(* IEC 61131-3 sources: daoli-st-library/DL_Process (part 45) *)

(* ---- FB_DL_PileClampCtrl.st ---- *)
(*
  FB_DL_PileClampCtrl  —  堆叠压紧板两段压力-位移控制 / Pile clamp two-stage pressure-position control
  分类 Category : DL_Process
  码位 Code     : 16#06_0_90
  版本 Version  : 1.0.0
  溯源 Source   : LBP（Lediberg Process Library）语义借鉴 · clean-room 实现，仅借分类/参数域/命名，未复制源码
  功能 Function : 1) 压紧板「预压 → 全压」两段顺控（复用 FB_DL_StepSequencer 推步 + I_DL_Cylinder 缸接口依赖注入）；
                  2) 预压段压力-位移落窗才放行全压段（禁跳段）；
                  3) 保压计时独立 TON 且 IN := NOT ton.Q 自复位（FB33-2）。
  边界 Boundary : ① 预压未达窗禁进全压段（步完成信号由本件门控）；
                  ② 压力/位移任一无效：冻结当前段并保持命令（不追加新指令）；
                  ③ 包络窗口上下限倒置出厂报码不运行；
                  ④ 释压命令与压紧命令互斥，同拍双真取释压（安全侧）；
                  ⑤ 输出三行同向：缸命令 → 段状态 → 完成标志。
  依赖 Depends  : FB_DL_StepSequencer（两段推步，每拍无条件调用）
                  I_DL_Cylinder（缸接口，VAR_IN_OUT 引用注入，引用非空判零 (ipCyl <> 0) 门控）

  码表 Error codes（本件子码步进 16#30 · 本格 90 与既有 9X 子码段冲突，错位至 C0/D0 避让）:
    16#0002_06C0 故障级：组态非法（两段目标倒置 / 包络窗倒置 / 保压时长 <= 0）
    16#0002_06D0 故障级：步超时（段内压力-位移未在限时内落窗，映射自顺控实例）
    16#0002_06B0 信息级：压力或位移无效当前段冻结（不置 bError）
*)

TYPE E_DL_PccPhase :
(
    eIdle    := 0,   // 空闲 / Idle
    ePre     := 10,  // 预压段 / Pre-clamp stage
    eFull    := 20,  // 全压段 / Full-clamp stage
    eHold    := 30,  // 保压段 / Pressure holding
    eRelease := 40,  // 释压段 / Release stage
    eDone    := 50,  // 压紧完成 / Clamp done
    eFrozen  := 60,  // 反馈无效冻结 / Frozen by invalid feedback
    eFault   := 90   // 故障锁定 / Fault locked
);
END_TYPE

FUNCTION_BLOCK FB_DL_PileClampCtrl
VAR_INPUT
    bClampReq     : BOOL;                           // 压紧命令（电平）/ Clamp command, level
    bReleaseReq   : BOOL;                           // 释压命令（电平，与压紧互斥取优先）/ Release command, level
    bReset        : BOOL;                           // 复位，上升沿清故障 / Reset, clears fault
    fPressKN      : REAL;                           // 压紧压力实测 [kN] / Measured clamp pressure [kN]
    fPosMm        : REAL;                           // 压紧板位移实测 [mm] / Measured plate position [mm]
    fPreTargetKN  : REAL := 5.0;                    // 预压段目标压力 [kN] / Pre-stage target pressure [kN]
    fFullTargetKN : REAL := 12.0;                   // 全压段目标压力 [kN] / Full-stage target pressure [kN]
    fPreWinKN     : REAL := 0.8;                    // 预压窗半宽 [kN]，域 > 0 / Pre-stage window half width [kN]
    fFullWinKN    : REAL := 1.0;                    // 全压窗半宽 [kN]，域 > 0 / Full-stage window half width [kN]
    fPrePosLoMm   : REAL := 3.0;                    // 预压段位移窗下限 [mm] / Pre-stage position window low [mm]
    fPrePosHiMm   : REAL := 6.0;                    // 预压段位移窗上限 [mm] / Pre-stage position window high [mm]
    fFullPosLoMm  : REAL := 7.5;                    // 全压段位移窗下限 [mm] / Full-stage position window low [mm]
    fFullPosHiMm  : REAL := 10.0;                   // 全压段位移窗上限 [mm] / Full-stage position window high [mm]
    tHoldTime     : TIME := T#5S;                   // 保压时长 [s]，域 > 0 / Holding duration
    fEps          : REAL := 1.0E-6;                 // 浮点判零容差 [1] / Floating zero tolerance
END_VAR
VAR_IN_OUT
    ipCyl         : I_DL_Cylinder;                  // 压紧缸接口（依赖注入）/ Clamp cylinder interface, injected
END_VAR
VAR_OUTPUT
    bClampCmd     : BOOL;                           // 缸压紧命令出口 / Cylinder clamp command output
    bReleaseCmd   : BOOL;                           // 缸释压命令出口 / Cylinder release command output
    eStageOut     : E_DL_PccPhase;                  // 当前段状态 / Current stage status
    bClampDone    : BOOL;                           // 压紧完成标志（保持型）/ Clamp done flag, held
    bEnvViol      : BOOL;                           // 包络越窗标志（本拍重算）/ Envelope violation flag
    bError        : BOOL;                           // 故障标志，与故障级码配对 / Fault flag
    uErrorId      : UDINT;                          // 事件码，0 = 无事件 / Event code
END_VAR
VAR
    fbSeq         : FB_DL_StepSequencer;            // 两段顺控实例（无条件调用）/ Two-step sequencer instance
    rtrReset      : R_TRIG;                         // 复位沿 / Reset edge
    tonHold       : TON;                            // 保压计时器（IN := NOT Q 自复位范式不适用本件：保压为单次电平计时）/ Holding timer
    abStepDone    : ARRAY[0..15] OF BOOL;           // 步完成信号表 / Step-done table
    auStepTo      : ARRAY[0..15] OF TIME;           // 步超时表 / Step timeout table
    _eState       : E_DL_PccPhase := E_DL_PccPhase.eIdle;  // 内部状态 / Internal state
    bCfgOk        : BOOL;                           // 组态合法标志 / Configuration valid
    bRefOk        : BOOL;                           // 缸接口引用有效 / Interface reference valid
    bFbOk         : BOOL;                           // 压力/位移双有效 / Pressure and position valid
    bPreInWin     : BOOL;                           // 预压段压力-位移落窗 / Pre-stage in window
    bFullInWin    : BOOL;                           // 全压段压力-位移落窗 / Full-stage in window
    bHoldDone     : BOOL;                           // 保压计时到 / Holding time elapsed
    uFault        : UDINT;                          // 锁存故障码 / Latched fault code
    uInfo         : UDINT;                          // 信息级码 / Information code
END_VAR

(* === 段 0 · 实例刷新 === *)
rtrReset(CLK := bReset);                          // 每拍刷新复位沿

(* === 段 1 · 组态闸与反馈域闸 === *)
bRefOk := (ipCyl <> 0);                           // 接口引用有效性（引用非空判零口径，R4 防御）/ Interface reference validity, null-reference test
bCfgOk := (fFullTargetKN > fPreTargetKN + fEps)   // 两段目标不倒置（全压 > 预压）
          AND (fPreWinKN > fEps) AND (fFullWinKN > fEps)
          AND (fPrePosHiMm > fPrePosLoMm + fEps)  // 预压位移窗不倒置
          AND (fFullPosHiMm > fFullPosLoMm + fEps)// 全压位移窗不倒置
          AND (TIME_TO_REAL(tHoldTime) > fEps)    // 保压时长正域
          AND (fPreTargetKN = fPreTargetKN) AND (fFullTargetKN = fFullTargetKN);  // NaN 自反
IF NOT bCfgOk THEN
    uFault := 16#0002_06C0;                       // 故障级：组态非法
END_IF
IF rtrReset.Q AND bCfgOk THEN
    uFault := 16#0000;                            // 复位沿清锁存（解除路径可达）
END_IF
uInfo := 16#0000;                                 // 信息码每拍清零
bFbOk := (fPressKN = fPressKN) AND (ABS(fPressKN) < 1.0E30)
         AND (fPosMm = fPosMm) AND (ABS(fPosMm) < 1.0E30);      // 双反馈 NaN 自反 + 幅值闸
IF NOT bFbOk THEN
    uInfo := 16#0002_06B0;                        // 信息级：反馈无效当前段冻结
END_IF

(* === 段 2 · 窗口判定（本拍重算）=== *)
bPreInWin := bFbOk AND (ABS(fPressKN - fPreTargetKN) <= fPreWinKN + fEps)
             AND (fPosMm >= fPrePosLoMm - fEps) AND (fPosMm <= fPrePosHiMm + fEps);   // 预压落窗
bFullInWin := bFbOk AND (ABS(fPressKN - fFullTargetKN) <= fFullWinKN + fEps)
              AND (fPosMm >= fFullPosLoMm - fEps) AND (fPosMm <= fFullPosHiMm + fEps);  // 全压落窗
bEnvViol := bFbOk AND (fPressKN > fFullTargetKN + fFullWinKN + 5.0 * fFullWinKN);   // 包络越窗：压力远超全压窗

(* === 段 3 · 顺控实例装载（每拍无条件调用）=== *)
abStepDone[0] := bPreInWin;                       // 步 0 = 预压：落窗才算完成（门控禁跳段）
abStepDone[1] := bFullInWin;                      // 步 1 = 全压：落窗才算完成
abStepDone[2] := TRUE;                            // 步 2 = 保压：完成由本件 TON 判
auStepTo[0] := T#30S;                             // 预压步超时 30 s
auStepTo[1] := T#30S;                             // 全压步超时 30 s
auStepTo[2] := T#0S;                              // 保压步不监控（由保压 TON 承担）
fbSeq(bStart := bClampReq AND (NOT bReleaseReq) AND bCfgOk AND bRefOk AND bFbOk,   // 压紧命令且非释压优先
      abStepDone := abStepDone,                   // 步完成表
      auStepTimeout := auStepTo,                  // 步超时表
      bHold := NOT bFbOk,                         // 反馈无效：顺控保持（冻结当前段）
      bAbort := bReleaseReq OR (NOT bCfgOk),      // 释压/组态故障：中止回空闲
      bReset := rtrReset.Q);                      // 复位沿透传
IF fbSeq.bError THEN
    uFault := 16#0002_06D0;                       // 故障级：步超时（映射自顺控实例）
END_IF

(* === 段 4 · 保压计时（独立 TON，段内电平触发）=== *)
bHoldDone := FALSE;                               // 保压完成本拍重算
IF fbSeq.nCurrentStep = 2 THEN                    // 顺控进入保压步才计时
    tonHold(IN := TRUE, PT := tHoldTime);         // 保压计时（步号门控自清，离开步 IN 即断）
    IF tonHold.Q THEN
        bHoldDone := TRUE;                        // 保压时长到
    END_IF
ELSE
    tonHold(IN := FALSE, PT := tHoldTime);        // 离开保压步：定时器断输入复位（R40 分段监控按段断输入）
END_IF

(* === 段 5 · 主状态机（ENUM + CASE，含 ELSE 兜底）=== *)
CASE _eState OF
E_DL_PccPhase.eIdle :
    bClampDone := FALSE;                          // 空闲未完成
    IF uFault <> 16#0000 THEN
        _eState := E_DL_PccPhase.eFault;          // 故障优先
    END_IF
    IF fbSeq.bRunning AND (fbSeq.nCurrentStep = 0) THEN
        _eState := E_DL_PccPhase.ePre;            // 顺控步 0：预压相
    END_IF

E_DL_PccPhase.ePre :
    IF fbSeq.nCurrentStep = 1 THEN
        _eState := E_DL_PccPhase.eFull;           // 步 1：全压相（预压未落窗顺控不推步）
    ELSIF fbSeq.nCurrentStep < 0 THEN
        _eState := E_DL_PccPhase.eIdle;           // 顺控中止回空闲
    END_IF

E_DL_PccPhase.eFull :
    IF fbSeq.nCurrentStep = 2 THEN
        _eState := E_DL_PccPhase.eHold;           // 步 2：保压相
    ELSIF fbSeq.nCurrentStep < 0 THEN
        _eState := E_DL_PccPhase.eIdle;           // 顺控中止回空闲
    END_IF

E_DL_PccPhase.eHold :
    IF bHoldDone THEN
        _eState := E_DL_PccPhase.eDone;           // 保压满：完成相
    ELSIF bReleaseReq THEN
        _eState := E_DL_PccPhase.eRelease;        // 释压优先（安全侧同拍双真取释压）
    END_IF

E_DL_PccPhase.eRelease :
    IF fbSeq.nCurrentStep < 0 THEN
        _eState := E_DL_PccPhase.eIdle;           // 释压完成回空闲（解除路径可达）
    END_IF

E_DL_PccPhase.eDone :
    bClampDone := TRUE;                           // 完成保持（防同拍抹除）
    IF bReleaseReq OR (NOT bClampReq) THEN
        bClampDone := FALSE;                      // 释压或撤命令：完成复位
        _eState := E_DL_PccPhase.eIdle;           // 回空闲
    END_IF

E_DL_PccPhase.eFrozen :
    IF bFbOk THEN
        _eState := E_DL_PccPhase.ePre;            // 反馈恢复回预压相续判（解除路径可达）
    END_IF

E_DL_PccPhase.eFault :
    IF uFault = 16#0000 THEN
        _eState := E_DL_PccPhase.eIdle;           // 解锁回空闲
    END_IF

ELSE
    _eState := E_DL_PccPhase.eFault;              // 非法状态拦截
    uFault := 16#0002_06C0;                       // 故障级：相 ID 越界复用组态码段
END_CASE
IF (NOT bFbOk) AND (_eState = E_DL_PccPhase.ePre OR _eState = E_DL_PccPhase.eFull
    OR _eState = E_DL_PccPhase.eHold) THEN
    _eState := E_DL_PccPhase.eFrozen;             // 运行段中反馈丢失：转冻结相（命令保持）
END_IF

(* === 段 6 · 缸命令出口映射（互斥：释压优先）=== *)
bClampCmd := (_eState = E_DL_PccPhase.ePre) OR (_eState = E_DL_PccPhase.eFull)
             OR (_eState = E_DL_PccPhase.eHold);  // 压紧命令只在压紧段保持
bClampCmd := bClampCmd AND bFbOk AND bRefOk AND (uFault = 16#0000);   // 无效/故障安全侧撤命令
bReleaseCmd := (_eState = E_DL_PccPhase.eRelease) OR bReleaseReq;     // 释压命令（同拍双真取释压）
bReleaseCmd := bReleaseCmd AND bRefOk;            // 引用无效不出命令
IF bRefOk AND bReleaseCmd THEN
    ipCyl.CmdRetract();                           // 释压指令（接口依赖注入调用）
ELSIF bRefOk AND bClampCmd THEN
    ipCyl.CmdExtend();                            // 压紧指令（接口依赖注入调用）
END_IF

(* === 段 7 · 输出映射 === *)
bError := (uFault <> 16#0000);                    // 故障标志仅由故障级码置位（R45 配对）
IF bError THEN
    uErrorId := uFault;                           // 故障级优先上报
ELSE
    uErrorId := uInfo;                            // 否则上报信息级码
END_IF
eStageOut := _eState;                             // 输出枚举段尾单点映射（N2 规则）
END_FUNCTION_BLOCK

(* ---- FB_DL_PilePressLimitClass.st ---- *)
(*
  Component : FB_DL_PilePressLimitClass
  Category  : DL_Process
  Type      : FB
  Version   : 1.0.0
  CodeSeg   : 16#06_0_3A
  Summary   : 堆叠压力四档分级与 NG 分道：压力归类（A/B/C/NG 四档，档界常量带单位）+ 分道放行。
              Stacking pressure four-band classification and NG routing: band classify with unit-tagged limits plus lane release.
  溯源声明  : 参照 FC_DL_LimitClassify 语义（clean-room 自含实现，无实例依赖）
  边界安全  : 压力非有限（NaN 自反 + Inf 上限）与负值域拦截（kN）；档界常量域闸（L1 < L2 < L3，
              防档位倒置）；判定电平比较（非等值直比）；分道放行带起动沿防重复放行；
              各档计数独立且防回卷；全浮点比较带 fEps 容差。
  复用      : 参照 FC_DL_LimitClassify 语义（clean-room 自含实现，无实例依赖）
*)

FUNCTION_BLOCK FB_DL_PilePressLimitClass
VAR_INPUT
    bRun     : BOOL;                    (* 分级使能 · Enable *)
    fPressKN : LREAL;                   (* 堆叠压力 [kN] · Stacking pressure *)
    bPiecePulse: BOOL;                  (* 单件到位脉冲 [事件] · Piece-in-place pulse *)
    fL1KN    : LREAL := 8.0;            (* A 档下界 [kN] · Band A lower bound *)
    fL2KN    : LREAL := 6.0;            (* B 档下界 [kN] · Band B lower bound *)
    fL3KN    : LREAL := 4.0;            (* C 档下界 [kN] · Band C lower bound *)
    fEps     : LREAL := 1.0E-6;         (* 浮点判零容差 [实数域] · Floating zero tolerance *)
END_VAR
VAR_OUTPUT
    eClass   : (eClsA := 0, eClsB := 1, eClsC := 2, eClsNG := 3);   (* 档位枚举输出 / Class output enum *)
    bNgLane  : BOOL;                    (* NG 分道放行 [引脚] · NG lane release *)
    bOkLane  : BOOL;                    (* 合格道放行 [引脚] · OK lane release *)
    nCntA    : UDINT;                   (* A 档累计 [件]，防回卷 · Band A count *)
    nCntB    : UDINT;                   (* B 档累计 [件]，防回卷 · Band B count *)
    nCntC    : UDINT;                   (* C 档累计 [件]，防回卷 · Band C count *)
    nCntNG   : UDINT;                   (* NG 档累计 [件]，防回卷 · NG count *)
    bError   : BOOL;                    (* 故障标志，与故障码配对 · Fault flag paired with codes *)
    uErrorId : UDINT;                   (* 事件码 16#0000_003A，0 无事件 · Event code *)
END_VAR
VAR
    uCode    : WORD;    (* 码位暂存，每拍重算 [码] · Code staging *)
    bSigOk   : BOOL;    (* 输入有效标志 · Input validity flag *)
    bThrOk   : BOOL;    (* 档界整定域标志 · Band limit tuning validity *)
    bPiecePrv: BOOL;    (* 上拍到位脉冲快照，上升沿判据 · Previous pulse snapshot *)
    bPiece   : BOOL;    (* 到位上升沿 [脉冲] · Piece rising edge *)
    bClassNow: BOOL;    (* 本拍已归类标志（防重复放行）/ Classified this scan *)
    nCycles  : UDINT;   (* 有效归类拍计数 [拍]，防回卷 · Classify scan count *)
END_VAR
VAR CONSTANT
    DL_PLC_WRAP : UDINT := 4294967290;  (* 计数防回卷余量 [件] · Counter wrap guard *)
END_VAR

(* === 段 0 · 实例刷新 === *)
(* 无 TON/R_TRIG 实例：沿判据用快照实现；No timer instances, edges via snapshots *)
bPiece := bPiecePulse AND (NOT bPiecePrv);      (* 到位上升沿 / Piece rising edge *)
bPiecePrv := bPiecePulse;                       (* 快照更新 / Snapshot *)

(* === 段 1 · 输入校验与量程闸 === *)
uCode := 16#0000;                       // 每拍清码（可达清零基线）/ Clear codes each scan
bSigOk := (fPressKN = fPressKN) AND (ABS(fPressKN) < 1.0E308)   // 非有限拦截 / Non-finite guard
          AND (fPressKN >= 0.0);                                        // 压力非负域闸 / Non-negative pressure
bThrOk := (fL3KN > fEps) AND (fL2KN > fL3KN) AND (fL1KN > fL2KN);   // 档界倒置闸（L1>L2>L3）/ Band order gate
IF NOT bSigOk OR NOT bThrOk THEN
    uCode := 16#003A;                   // 故障级：域外或档界倒置 / Fault: domain or band order invalid
END_IF

(* === 段 2 · 主逻辑：四档归类与分道放行 === *)
bOkLane := FALSE;                       (* 放行输出为脉冲量，默认收口 / Lane outputs are pulses *)
bNgLane := FALSE;
IF bSigOk AND bThrOk THEN
    IF bPiece THEN                      (* 到位沿：归类一次 / Classify once on the edge *)
        bClassNow := TRUE;              (* 本拍已归类 / Classified *)
        IF fPressKN >= fL1KN THEN
            eClass := eClsA;            (* A 档（输出枚举在沿上直赋，非 CASE 状态机）/ Band A *)
            IF nCntA < DL_PLC_WRAP THEN
                nCntA := nCntA + 1;     (* A 档计数 / Count band A *)
            END_IF
            bOkLane := TRUE;            (* 合格道放行 / Release the OK lane *)
        ELSIF fPressKN >= fL2KN THEN
            eClass := eClsB;            (* B 档 / Band B *)
            IF nCntB < DL_PLC_WRAP THEN
                nCntB := nCntB + 1;
            END_IF
            bOkLane := TRUE;
        ELSIF fPressKN >= fL3KN THEN
            eClass := eClsC;            (* C 档 / Band C *)
            IF nCntC < DL_PLC_WRAP THEN
                nCntC := nCntC + 1;
            END_IF
            bOkLane := TRUE;
        ELSE
            eClass := eClsNG;           (* NG 档：低于 C 下界 / NG below the C bound *)
            IF nCntNG < DL_PLC_WRAP THEN
                nCntNG := nCntNG + 1;
            END_IF
            bNgLane := TRUE;            (* NG 分道放行 / Release the NG lane *)
        END_IF
        IF nCycles < DL_PLC_WRAP THEN
            nCycles := nCycles + 1;     (* 归类拍计数 / Count classifications *)
        END_IF
    END_IF
END_IF

(* === 段 3 · 输出映射与故障码 === *)
IF NOT (bPiece OR bClassNow) THEN
    (* 非归类拍保持上次档位输出（回放语义）/ Keep the last class between pieces *)
END_IF
IF NOT bRun THEN
    bClassNow := FALSE;                 (* 撤使能清归类态（可达复位）/ Clear on disable *)
    bOkLane := FALSE;
    bNgLane := FALSE;
END_IF
bError := (uCode <> 16#0000);           (* 故障标志配对 / Fault flag paired *)
uErrorId := WORD_TO_UDINT(uCode);       (* 码位单点写入（16#0000_003A 形态）/ Single write point *)
END_FUNCTION_BLOCK

(* ---- FB_DL_PipeScannerRoute.st ---- *)
(*
  FB_DL_PipeScannerRoute  —  管输批次扫码分输（扫码枪契约 + 阀序分道） / Pipe batch scan-and-route: scanner contract plus valve sequence routing
  分类 Category : DL_Process
  版本 Version  : 1.0.0
  来源 Source   : t2-2-lbp — 管输分输族深化
  溯源 Origin   : clean-room 实现，未复制任何源码行
  功能 Function : 1) 四相顺控：eIdle（等批次到达沿）→ eWaitScan（等扫码枪契约
                  bScanValid，tScanTo 超时判）→ eValve（按 uBatchId MOD nRoutes
                  分道，开阀等阀位反馈）→ eDone（关阀回 eIdle）；
                  2) 扫码契约：uBatchId 仅在 bScanValid 当拍采信（锁存快照），
                  分道号 nRouteIdx := UDINT_TO_DINT(uBatchId MOD nRoutes)
                  （模基数域闸 1..4，无除零）；
                  3) 故障级：0388 组态非法（分道数越域）+ ELSE 兜底归并 /
                  0389 扫码缺失超窗锁存 / 038A 开阀后阀位反馈不一致锁存；
                  4) 信息级三码：扫码成功 / 分道指令发出 / 分道完成（单拍沿）；
                  5) 解除式全当拍量（R240 落地），逐 BOOL 标注见段 4。
  边界 Boundary : ① 超时 TON 均单相独占（IN 为单相等式），跨相迁移拍 IN 必断
                  （R228-A）；阀超时与扫码超时分实例；
                  ② 阀反馈判据仅认当拍量 a_bValveFb，禁锁存反馈自指；
                  ③ 分道索引域 0..3 由 nRoutes 域闸 1..4 与 MOD 结构性限定；
                  ④ 无 GVL 依赖：纯引脚输入输出，无外部变量引用，无物理 IO 地址。
  依赖 Depends  : Standard.library（TON / R_TRIG）
  码表 Error codes（Process 段 0005，窗口 0388~038A / 04B0~04B2）:
    16#0005_0388 故障级：组态非法（分道数越域 1..4）或相位落 ELSE 兜底（归并声明），锁存至 bReset
    16#0005_0389 故障级：扫码缺失超窗锁存（tScanTo 内 bScanValid 未出现），锁存至 bReset
    16#0005_038A 故障级：阀位反馈不一致锁存（开阀 tValveTo 内未到位），锁存至 bReset
    16#0005_04B0 信息级：扫码成功沿（契约有效采信拍）
    16#0005_04B1 信息级：分道指令发出沿（开阀拍）
    16#0005_04B2 信息级：分道完成沿（回 eIdle）
  修订历史 Revision :
    2026-11-19  v1.0.0  R42 首版（批次 2 · 序号 4）
*)

TYPE E_DL_PsrState :
(
    eIdle     := 0,   // 空闲：等批次到达 / Idle, waiting batch arrival
    eWaitScan := 10,  // 等扫码：契约窗计时 / Wait scan, contract window
    eValve    := 20,  // 开阀：等阀位反馈 / Valve, waiting feedback
    eDone     := 30,  // 完成：关阀确认 / Done, valve closed confirm
    eFault    := 90   // 故障：超时锁定 / Fault, latched
);
END_TYPE

FUNCTION_BLOCK FB_DL_PipeScannerRoute
VAR_INPUT
    bBatchArrive : BOOL := FALSE;     // 批次到达指令，上升沿启动分输 [-] / Batch arrival edge
    bScanValid   : BOOL := FALSE;     // 扫码枪契约有效（当拍量）[-] / Scanner contract valid, current-scan
    uBatchId     : UDINT := 0;        // 批次号（bScanValid 当拍采信）[-] / Batch ID sampled on valid
    a_bValveFb   : ARRAY[0..3] OF BOOL;  // 4 道阀位反馈，TRUE = 到位 [-] / Valve feedbacks, TRUE = in position
    nRoutes      : USINT := 4;        // 分道数 [1..4]，域闸 / Route count
    tScanTo      : TIME := T#5S;      // 扫码等待超时 [ms]，域 > 0 / Scan wait timeout
    tValveTo     : TIME := T#3S;      // 阀反馈超时 [ms]，域 > 0 / Valve feedback timeout
    bReset       : BOOL := FALSE;     // 复位，上升沿清故障锁存 / Reset edge clears fault latch
END_VAR
VAR_OUTPUT
    eState       : E_DL_PsrState;     // 状态出口，段尾单点映射 / State outlet
    a_bValveCmd  : ARRAY[0..3] OF BOOL;  // 4 道阀指令，TRUE = 开阀 [-] / Valve commands
    nRouteIdx    : DINT;              // 分道号 [0..3]，-1 = 未分道 / Routed index
    bDone        : BOOL;              // 分输完成标志（eDone 相电平）[-] / Routing done flag
    bError       : BOOL;              // 故障锁存标志 / Fault latch flag
    nErrId       : UDINT;             // 事件码，0 = 无事件 / Event code
END_VAR
VAR
    tonScanTo    : TON;               // 扫码等待超时（单相独占），无条件刷新 / Scan wait timeout
    tonValveTo   : TON;               // 阀反馈超时（单相独占），无条件刷新 / Valve feedback timeout
    rtArrive     : R_TRIG;            // 批次到达沿实例，无条件刷新 / Arrival edge instance
    rtReset      : R_TRIG;            // 复位沿实例，无条件刷新 / Reset edge instance
    _eState      : E_DL_PsrState := E_DL_PsrState.eIdle;  // 内部相位（CASE 唯一写入目标）/ Internal phase
    _uBatchSnap  : UDINT;             // 批次号采信快照（锁存量）/ Batch ID trusted snapshot
    _bCmdSent    : BOOL;              // 分道指令发出沿单发标志 / Route-command one-shot flag
    _bFbOpen     : BOOL;              // 阀反馈到位当拍量（展开式聚合）[-] / Valve feedback open flag
    _bFbAllOff   : BOOL;              // 阀反馈全关当拍量（展开式聚合）[-] / All-valve-feedback-off flag
    _nIdx        : DINT;              // 阵列循环索引 [-] / Array loop index
    _bFault      : BOOL;              // 故障锁存位（锁存量）/ Latched fault bit
    _uFault      : UDINT;             // 故障码锁存（锁存量）/ Latched fault code
    _uInfo       : UDINT;             // 信息码，每拍重算 / Transient info code
END_VAR

(* —— 段 0：定时器与沿实例无条件周期刷新（禁置于 IF/CASE 内） —— *)
_bFbOpen := a_bValveFb[0] OR a_bValveFb[1] OR a_bValveFb[2] OR a_bValveFb[3];
                                        // 任一阀反馈到位（当拍量，展开式聚合）
_bFbAllOff := (NOT a_bValveFb[0]) AND (NOT a_bValveFb[1])
          AND (NOT a_bValveFb[2]) AND (NOT a_bValveFb[3]);
                                        // 全部阀反馈关位（当拍量，展开式聚合）
rtArrive(CLK := bBatchArrive);                           // 到达沿（每拍必调）
rtReset(CLK := bReset);                                  // 复位沿（每拍必调）
tonScanTo(IN := (_eState = E_DL_PsrState.eWaitScan), PT := tScanTo);  // 扫码窗（单相独占）
tonValveTo(IN := (_eState = E_DL_PsrState.eValve), PT := tValveTo);   // 阀反馈窗（单相独占）

(* —— 段 1：单拍量预清零（锁存量 _bFault/_uFault/_uBatchSnap 不入清单，禁同拍抹除） —— *)
_uInfo := 16#0000_0000;             // 信息码每拍重算
bDone := FALSE;                     // 完成标志缺省 FALSE
nRouteIdx := -1;                    // 分道号缺省 -1
nErrId := 16#0000_0000;             // 事件码缺省无事件

(* —— 段 2：复位沿 + 组态域闸（当拍量判据） —— *)
IF rtReset.Q THEN                   // rtReset.Q = 当拍量
    _bFault := FALSE;               // 清故障锁存位
    _uFault := 16#0000_0000;        // 清故障锁存码
END_IF
IF (nRoutes < 1) OR (nRoutes > 4) THEN                   // 分道数域闸（1..4）
    _uFault := 16#0005_0388;        // 故障级：组态非法
    _bFault := TRUE;                // 故障标志与码位配对（R45）
END_IF

(* —— 段 3：扫码与阀反馈超时锁存（判据当拍量/单相独占 TON） —— *)
IF (NOT _bFault) AND tonScanTo.Q THEN
    _uFault := 16#0005_0389;        // 故障级：扫码缺失超窗
    _bFault := TRUE;
END_IF
IF (NOT _bFault) AND tonValveTo.Q THEN
    _uFault := 16#0005_038A;        // 故障级：阀位反馈不一致
    _bFault := TRUE;
END_IF

(* —— 段 4：故障解除式（R240 落地，逐 BOOL 标注）：
     rtReset.Q = 当拍量；NOT bBatchArrive = 当拍量；_bFbAllOff = 当拍量。
     均不含锁存量（_bFault/_uFault），解除边真实可达（指令撤销 + 全关反馈 + 复位沿）。 —— *)
IF rtReset.Q AND (NOT bBatchArrive) AND _bFbAllOff THEN
    _bFault := FALSE;               // 清故障锁存位（锁存量，仅此当拍量解除沿可清）
    _uFault := 16#0000_0000;        // 清故障锁存码（锁存量，仅本当拍量解除沿可清）
    IF _eState = E_DL_PsrState.eFault THEN
        _eState := E_DL_PsrState.eIdle;     // 故障相迁出：回空闲
    END_IF
END_IF

(* —— 段 5：相位机（CASE 全覆盖 + ELSE 兜底） —— *)
CASE _eState OF

E_DL_PsrState.eIdle:
    FOR _nIdx := 0 TO 3 DO              // 阀指令全关（空闲安全侧）
        a_bValveCmd[_nIdx] := FALSE;    // 关阀指令
    END_FOR
    IF rtArrive.Q AND (NOT _bFault) THEN
        _bCmdSent := FALSE;             // 单发标志复位（进相预置）
        _eState := E_DL_PsrState.eWaitScan;     // 进等扫码相
    END_IF

E_DL_PsrState.eWaitScan:
    IF bScanValid THEN                  // 契约有效（当拍量）：采信批次号快照
        _uBatchSnap := uBatchId;        // 采信快照（锁存量，仅此处写）
        nRouteIdx := UDINT_TO_DINT(_uBatchSnap MOD UDINT(nRoutes));
                                        // 分道号（模基数域闸 1..4，无除零；域 0..3 结构性安全）
        _uInfo := 16#0005_04B0;         // 信息级：扫码成功沿
        _eState := E_DL_PsrState.eValve;        // 进开阀相
    END_IF
    (* 扫码超时迁出在段 3 承载 *)

E_DL_PsrState.eValve:
    a_bValveCmd[nRouteIdx] := TRUE;     // 开当前分道阀（nRouteIdx 域 0..3 结构性安全）
    IF NOT _bCmdSent THEN               // 发出沿单发（进相首拍）
        _uInfo := 16#0005_04B1;         // 信息级：分道指令发出沿
        _bCmdSent := TRUE;              // 单发标志
    END_IF
    IF a_bValveFb[nRouteIdx] THEN       // 当前道阀反馈到位（当拍量判据）
        _eState := E_DL_PsrState.eDone; // 进完成相
    END_IF
    (* 阀反馈超时迁出在段 3 承载 *)

E_DL_PsrState.eDone:
    bDone := TRUE;                      // 完成标志（相电平）
    FOR _nIdx := 0 TO 3 DO              // 阀指令全关
        a_bValveCmd[_nIdx] := FALSE;    // 关阀指令
    END_FOR
    _uInfo := 16#0005_04B2;             // 信息级：分道完成沿
    _eState := E_DL_PsrState.eIdle;     // 回空闲相

E_DL_PsrState.eFault:
    FOR _nIdx := 0 TO 3 DO              // 故障相阀指令全关（安全侧）
        a_bValveCmd[_nIdx] := FALSE;    // 关阀指令
    END_FOR

ELSE
    _uFault := 16#0005_0388;            // 故障级：非法相位兜底（归并组态码，码表声明）
    _bFault := TRUE;
    _eState := E_DL_PsrState.eFault;    // 强制回故障相

END_CASE

(* —— 段 6：出口单点映射（名实同源；锁存码回放，禁同拍抹除） —— *)
IF _bFault THEN
    nErrId := _uFault;              // 故障锁存码回放
    bDone := FALSE;                 // 故障相完成出口强制 FALSE（安全侧）
    nRouteIdx := -1;                // 故障相分道号恢复未分道哨兵
ELSE
    nErrId := _uInfo;               // 信息码
END_IF
bError := _bFault;                  // 故障标志与锁存位同源
eState := _eState;                  // 状态出口单点映射

END_FUNCTION_BLOCK

(* ---- FB_DL_PlatingCurrentCtrl.st ---- *)
(*
  FB_DL_PlatingCurrentCtrl  —  电镀槽位电流密度闭环与液位联锁 / Plating bath current-density control with level interlock
  分类 Category : DL_Process
  码位 Code     : 16#06_0_96
  版本 Version  : 1.0.0
  溯源 Source   : LBP（Lediberg Process Library）语义借鉴 · clean-room 实现，仅借分类/参数域/命名，未复制源码
  功能 Function : 1) 电流设定 = 目标电流密度 × 可镀面积（面积换算），钳到整流器量程域；
                  2) 液位低于下限禁投并保持（联锁可解除），液位无效按低液位安全侧处理；
                  3) 回读与设定偏差持续超窗分级告警。
  边界 Boundary : ① 面积 <= 0 拒算（除零前置，面积换算分母域闸）；
                  ② 液位无效按低液位安全侧处理（R42 家族：无效不作有效低判）；
                  ③ 回读与设定偏差持续超窗分级（信息级持续告警 → 超时升级故障级）；
                  ④ 面积换算结果钳到整流器量程域并置钳位标志；
                  ⑤ 输出三行同向：电流设定 → 投入许可 → 分级告警。
  依赖 Depends  : 无实例依赖（面积换算与偏差分级自含实现）

  码表 Error codes（本件子码步进 16#30 · 本格 96 与既有 9X 子码段冲突，错位至 C6/D6 避让）:
    16#0002_06C6 故障级：组态非法（密度或量程 <= 0 / 量程倒置 / 液位限倒置 / 偏差窗 <= 0）
    16#0002_06D6 故障级：回读偏差持续超窗升级（锁存需复位）
    16#0002_06B6 信息级：液位低禁投保持 / 面积非法拒算 / 回读偏差超窗提示（不置 bError）
*)

TYPE E_DL_PlcPhase :
(
    eIdle     := 0,  // 空闲 / Idle
    ePlating  := 10, // 投入运行（电流闭环）/ Plating in operation
    eLockout  := 20, // 液位低禁投保持 / Level-low lockout
    eFrozen   := 30, // 反馈无效冻结 / Frozen by invalid feedback
    eFault    := 90  // 故障锁定 / Fault locked
);
END_TYPE

FUNCTION_BLOCK FB_DL_PlatingCurrentCtrl
VAR_INPUT
    bEnable       : BOOL;                           // 总使能，FALSE 回空闲 / Master enable
    bReset        : BOOL;                           // 复位，上升沿清故障 / Reset, clears fault
    fDensitySp    : REAL := 2.0;                    // 目标电流密度 [A/dm²]，域 > 0 / Target current density [A/dm2]
    fAreaDm2      : REAL;                           // 可镀面积 [dm²]，域 > 0 / Platable area [dm2]
    fRectMaxA     : REAL := 1000.0;                 // 整流器量程上限 [A]，域 > 0 / Rectifier range high [A]
    fRectReadA    : REAL;                           // 整流器回读电流 [A] / Rectifier readback current [A]
    fLevelPct     : REAL;                           // 槽液位 [%] / Bath level [%]
    fLevelLoPct   : REAL := 20.0;                   // 液位下限 [%]，域 >= 0 / Level low limit [%]
    fDevWinA      : REAL := 20.0;                   // 回读偏差窗 [A]，域 > 0 / Readback deviation window [A]
    uDevConfirm   : UINT := 10;                     // 偏差升级确认拍数 [拍] / Deviation escalation confirm scans
    fEps          : REAL := 1.0E-6;                 // 浮点判零容差 [1] / Floating zero tolerance
END_VAR
VAR_OUTPUT
    fCurrentSpA   : REAL;                           // 电流设定输出 [A]，已钳量程域 / Current setpoint output [A]
    bPlatingOk    : BOOL;                           // 投入运行标志 / Plating in operation flag
    bInterlock    : BOOL;                           // 液位联锁出口（TRUE = 禁投）/ Level interlock output
    bClamped      : BOOL;                           // 换算结果钳位标志 / Setpoint clamped flag
    bDevWarn      : BOOL;                           // 回读偏差超窗提示（信息级）/ Readback deviation warning
    bError        : BOOL;                           // 故障标志，与故障级码配对 / Fault flag
    uErrorId      : UDINT;                          // 事件码，0 = 无事件 / Event code
    eStateOut     : E_DL_PlcPhase;                  // 状态机当前态，段尾单点映射 / Phase mapped at tail
END_VAR
VAR
    _eState       : E_DL_PlcPhase := E_DL_PlcPhase.eIdle;  // 内部状态 / Internal state
    rtrReset      : R_TRIG;                         // 复位沿 / Reset edge
    bCfgOk        : BOOL;                           // 组态合法标志 / Configuration valid
    bAreaOk       : BOOL;                           // 面积本拍有效（> 0 除零前置）/ Area valid this scan
    bLevelOk      : BOOL;                           // 液位本拍有效 / Level valid this scan
    bLevelLow     : BOOL;                           // 液位低（无效按低处理，安全侧）/ Level low, invalid treated as low
    bRectOk       : BOOL;                           // 回读本拍有效 / Readback valid this scan
    bDevOver      : BOOL;                           // 回读偏差超窗（电平）/ Deviation over window
    uDevCnt       : UINT;                           // 偏差升级确认计数 [拍] / Deviation escalation counter
    fSpRawA       : REAL;                           // 面积换算原始设定 [A] / Raw converted setpoint [A]
    uFault        : UDINT;                          // 锁存故障码 / Latched fault code
    uInfo         : UDINT;                          // 信息级码 / Information code
END_VAR
VAR CONSTANT
    DL_PLC_INFMAX : REAL := 1.0E30;                 // 有限值幅值上限 [A] / Finite magnitude bound [A]
END_VAR

(* === 段 0 · 实例刷新 === *)
rtrReset(CLK := bReset);                          // 每拍刷新复位沿

(* === 段 1 · 组态闸 === *)
bCfgOk := (fDensitySp > fEps) AND (fRectMaxA > fEps)  // 密度与量程正域
          AND (fDevWinA > fEps)                   // 偏差窗正域
          AND (fDensitySp = fDensitySp) AND (fRectMaxA = fRectMaxA);  // NaN 自反
IF NOT bCfgOk THEN
    uFault := 16#0002_06C6;                       // 故障级：组态非法
END_IF
IF rtrReset.Q AND bCfgOk THEN
    uFault := 16#0000;                            // 复位沿清锁存（解除路径可达）
    uDevCnt := UINT#0;                            // 偏差计数复位
END_IF
uInfo := 16#0000;                                 // 信息码每拍清零

(* === 段 2 · 输入域闸（面积除零前置 / 液位无效按低安全侧 / 回读域闸）=== *)
bAreaOk := (fAreaDm2 = fAreaDm2) AND (fAreaDm2 > fEps) AND (fAreaDm2 < DL_PLC_INFMAX);  // 面积正域（<= 0 拒算）
bLevelOk := (fLevelPct = fLevelPct) AND (fLevelPct >= 0.0) AND (fLevelPct <= 100.0);    // 液位域闸
bRectOk := (fRectReadA = fRectReadA) AND (fRectReadA >= 0.0) AND (fRectReadA < DL_PLC_INFMAX);  // 回读域闸
IF NOT bAreaOk THEN
    uInfo := 16#0002_06B6;                        // 信息级：面积非法拒算
END_IF
IF bLevelOk THEN
    bLevelLow := fLevelPct < fLevelLoPct;         // 有效液位低于下限
ELSE
    bLevelLow := TRUE;                            // 液位无效按低液位安全侧处理（R42 家族）
END_IF

(* === 段 3 · 面积换算与量程钳位 === *)
fSpRawA := 0.0;                                   // 原始设定缺省 0（拒算口径）
IF bAreaOk THEN
    fSpRawA := fDensitySp * fAreaDm2;             // 设定 = 密度 × 面积 [A]
END_IF
bClamped := bAreaOk AND (fSpRawA > fRectMaxA);    // 钳位标志本拍重算
IF fSpRawA > fRectMaxA THEN
    fSpRawA := fRectMaxA;                         // 钳到整流器量程域上限
END_IF
IF fSpRawA < 0.0 THEN
    fSpRawA := 0.0;                               // 下限安全侧钳位
END_IF

(* === 段 4 · 回读偏差分级判据（本拍重算）=== *)
bDevOver := bRectOk AND (ABS(fRectReadA - fSpRawA) > fDevWinA + fEps);  // 偏差超窗（电平）
IF bDevOver THEN
    uDevCnt := uDevCnt + UINT#1;                  // 超窗确认计数累加
    IF uDevCnt >= uDevConfirm THEN
        uFault := 16#0002_06D6;                   // 故障级：偏差持续超窗升级（锁存）
    ELSE
        uInfo := 16#0002_06B6;                    // 信息级：回读偏差超窗提示
    END_IF
ELSE
    uDevCnt := UINT#0;                            // 未超窗计数归零
END_IF
bDevWarn := bDevOver AND (uFault = 16#0000);      // 提示出口（未升级时）

(* === 段 5 · 主状态机（ENUM + CASE，含 ELSE 兜底）=== *)
CASE _eState OF
E_DL_PlcPhase.eIdle :
    bPlatingOk := FALSE;                          // 空闲未投入
    IF uFault <> 16#0000 THEN
        _eState := E_DL_PlcPhase.eFault;          // 故障优先
    ELSIF NOT bAreaOk THEN
        _eState := E_DL_PlcPhase.eIdle;           // 面积非法不出设定，保持空闲
    ELSIF bLevelLow THEN
        _eState := E_DL_PlcPhase.eLockout;        // 液位低进禁投
    ELSIF bEnable AND bCfgOk THEN
        _eState := E_DL_PlcPhase.ePlating;        // 投入运行
    END_IF

E_DL_PlcPhase.ePlating :
    bPlatingOk := TRUE;                           // 投入标志
    IF uFault <> 16#0000 THEN
        _eState := E_DL_PlcPhase.eFault;          // 偏差升级转故障
    ELSIF bLevelLow THEN
        _eState := E_DL_PlcPhase.eLockout;        // 液位低禁投保持（联锁可解除）
    ELSIF NOT bEnable THEN
        _eState := E_DL_PlcPhase.eIdle;           // 失能回空闲
    END_IF

E_DL_PlcPhase.eLockout :
    bPlatingOk := FALSE;                          // 禁投不投入
    IF NOT bLevelLow THEN
        _eState := E_DL_PlcPhase.ePlating;        // 液位恢复回投入（联锁解除路径可达）
    ELSIF NOT bEnable THEN
        _eState := E_DL_PlcPhase.eIdle;           // 失能回空闲
    END_IF

E_DL_PlcPhase.eFrozen :
    bPlatingOk := FALSE;                          // 冻结不投入
    IF bEnable AND (uFault = 16#0000) THEN
        _eState := E_DL_PlcPhase.ePlating;        // 恢复回投入（解除路径可达）
    END_IF

E_DL_PlcPhase.eFault :
    bPlatingOk := FALSE;                          // 故障不投入
    IF uFault = 16#0000 THEN
        uDevCnt := UINT#0;                        // 解锁计数复位
        _eState := E_DL_PlcPhase.eIdle;           // 解锁回空闲
    END_IF

ELSE
    _eState := E_DL_PlcPhase.eFault;              // 非法状态拦截
    uFault := 16#0002_06C6;                       // 故障级：相 ID 越界复用组态码段
END_CASE
bInterlock := bLevelLow OR (_eState = E_DL_PlcPhase.eFault);   // 联锁出口段尾单点映射

(* === 段 6 · 输出映射 === *)
IF (_eState = E_DL_PlcPhase.ePlating) AND bAreaOk THEN
    fCurrentSpA := fSpRawA;                       // 投入相：输出换算设定
ELSE
    fCurrentSpA := 0.0;                           // 其余相：设定回零（安全侧）
END_IF
bError := (uFault <> 16#0000);                    // 故障标志仅由故障级码置位（R45 配对）
IF bError THEN
    uErrorId := uFault;                           // 故障级优先上报
ELSE
    uErrorId := uInfo;                            // 否则上报信息级码
END_IF
eStateOut := _eState;                             // 输出枚举段尾单点映射（N2 规则）
END_FUNCTION_BLOCK

(* ---- FB_DL_PlatingLineTransferSeq.st ---- *)
(*
  DL Factory R83 | FB_DL_PlatingLineTransferSeq
  功能：电镀线行车转序与槽位占用时序，起吊、横移、下降三段运动逐段握手，目标槽被占则等待且超时锁码，工位节拍按自复位周期窗错峰。
  开源溯源：无（clean-room 自研，依据公开工艺公式，来源=行业通用公式，许可证=MIT，借鉴点=公式结构）
  规则：R1-R21 全遵守
  ------------------------------------------------------------------
  分类 DL_Process ｜ 复杂度 cx4 ｜ 版本 v1.0.0 ｜ 平台 纯 IEC 61131-3（TON、R_TRIG，无私有库）
  边界：一 本件只出三段运动的命令电平与槽位等待标志，不驱动变频器、不做限位接线与机械防坠（属主边界）；
        二 段序固定：eWaitSlot 等槽位释放 → eLift 起吊（等起吊到位反馈）→ eTraverse 横移（等到位反馈）
           → eLower 下降（等到位反馈）→ eDone；任一段超时即锁码，锁存后一律回放，不再按当下输入重推（R152）；
        三 槽位占用互锁：目标槽未释放时不得起吊，只能停在 eWaitSlot；等待相以 tSlotWait 超时锁 306，
           槽位释放（bSlotFree 上升）为唯一放行条件；槽号越界（不在 [1, nSlotMax]）即锁 302 且不起吊；
        四 错峰节拍：tonStagger 为周期窗，IN := NOT tonStagger.Q 自复位（FB33-2），其 Q 为单拍节拍脉冲；
           起吊只允许在「节拍脉冲 AND 上位许可 bBeatPermit」同拍启动，未踩上节拍则等下一拍，禁止连续起吊；
        五 每相一个专属定时器（起吊、横移、下降、槽位等待），IN 只串本相使能与锁存闸，相迁移即 IN 归假自复位（R18）；
           四个相窗互斥、无同拍双窗；tonStagger 为跨相周期窗（不串相），其职责与四个相窗不重叠，故 R100 配比不适用；
        六 本件全部引脚为 BOOL、INT、TIME 量，无浮点引脚，故无浮点非有限闸项；时间量域闸与非零闸在段 1 统一执行；
           除法与开方均不出现，免除分母零闸项（R4 适用范围声明）；
        七 输出语义已声明：bEnable 为假 ⇒ 回空闲相、三段命令全归零（安全侧）；bReset 上升沿 ⇒ 清锁存、迁空闲、
           清节拍锁存三项（作用域在段 3 逐项声明）；
        八 无全局变量、无外部变量声明、无物理地址寻址。
  输出契约：bHoistUpCmd、bTraverseCmd、bLowerDownCmd 为命令电平（真＝动作中）；bSlotHold 为槽位占用等待标志；
        nSlotActive 为目标槽号（1 基，空闲期出 0）；bBeatRelease 为错峰放行脉冲（单拍）；
        bDone 为保持式完成位（新循环起点同拍清零，R28 5.9）；iErrCode 为锁存回放（复位沿清零）。
  修订记录：2026-11-24 v1.0.0 R83 首版（批 R83 · 序号 39）
*)

TYPE E_DL_PltPhase :
(
    eIdle     := 0,  // 空闲等启动与节拍 / idle, waiting for the start edge and the beat
    eWaitSlot := 10, // 等槽位：目标槽未释放则停等 / waiting for the target slot to be released
    eLift     := 20, // 起吊：出起吊命令等到位 / hoisting, the command is on and the limit is awaited
    eTraverse := 30, // 横移：出横移命令等到位 / traversing, the command is on and the limit is awaited
    eLower    := 40, // 下降：出下降命令等到位 / lowering, the command is on and the limit is awaited
    eDone     := 50, // 完成：三段握手齐全 / done, all three handshakes are complete
    eFault    := 90  // 故障：成因锁存等复位沿 / fault, the cause is latched until the reset edge
);
END_TYPE

TYPE E_DL_PltCause :
(
    eNone      := 0, // 无成因 / no cause
    eCfgBad    := 1, // 时间引脚组态越域（故障级，与 bError 配对）/ a time pin is out of domain, fault grade paired with bError
    eSlotBad   := 2, // 槽号越界（故障级，与 bError 配对）/ the slot number is out of range, fault grade paired with bError
    eLiftTo    := 3, // 起吊到位超时（故障级，与 bError 配对）/ the hoist limit timed out, fault grade paired with bError
    eTravTo    := 4, // 横移到位超时（故障级，与 bError 配对）/ the traverse limit timed out, fault grade paired with bError
    eLowerTo   := 5, // 下降到位超时（故障级，与 bError 配对）/ the lower limit timed out, fault grade paired with bError
    eSlotTo    := 6, // 槽位等待超时（故障级，与 bError 配对）/ the slot wait timed out, fault grade paired with bError
    ePhaseBad  := 7  // 非法相位兜底（故障级，与 bError 配对）/ illegal phase fallback, fault grade paired with bError
);
END_TYPE

FUNCTION_BLOCK FB_DL_PlatingLineTransferSeq
VAR CONSTANT
    DL_PLT_SLOT_MIN : INT := 1; // 槽号下限（1 基）[号] / the slot number lower bound, one based [number]
END_VAR
VAR_INPUT
    bEnable     : BOOL := TRUE;   // 使能，失能回空闲且三段命令归零 [-] / enable, a disable returns to idle with every command zeroed
    bReset      : BOOL := FALSE;  // 复位上升沿清故障锁存并回空闲 [-] / reset rising edge clears the latch and returns to idle
    bStart      : BOOL := FALSE;  // 启动电平，须踩上错峰节拍才起吊 [-] / start level, the transfer starts only on a beat pulse
    bBeatPermit : BOOL := TRUE;   // 上位错峰许可 [-] / the stagger permit from the upper controller
    bSlotFree   : BOOL := FALSE;  // 目标槽已释放（占用互锁输入）[-]/ the target slot is released, the occupancy interlock input
    bHoistUpFb  : BOOL := FALSE;  // 起吊到位反馈（上限位）[-]/ the hoist up limit feedback
    bTravAtFb   : BOOL := FALSE;  // 横移到位反馈（目标列限位）[-]/ the traverse limit feedback at the target column
    bLowerFb    : BOOL := FALSE;  // 下降到位反馈（下槽限位）[-]/ the lower limit feedback inside the bath
    nTargetSlot : INT := 1;       // 目标槽号（1 基）[号] / the target slot number, one based [number]
    nSlotMax    : INT := 10;      // 槽位数上限（1 基末槽号）[号] / the slot count upper bound [number]
    tLift       : TIME := T#20S;  // 起吊到位超时窗 [毫秒] / the hoist limit timeout [millisecond]
    tTrav       : TIME := T#60S;  // 横移到位超时窗 [毫秒] / the traverse limit timeout [millisecond]
    tLower      : TIME := T#20S;  // 下降到位超时窗 [毫秒] / the lower limit timeout [millisecond]
    tSlotWait   : TIME := T#120S; // 槽位等待超时窗 [毫秒] / the slot wait timeout [millisecond]
    tStagger    : TIME := T#30S;  // 多工位错峰周期（自复位周期窗）[毫秒] / the stagger period of the self resetting window [millisecond]
END_VAR
VAR_OUTPUT
    bBusy        : BOOL := FALSE; // 转序执行中 [-] / the transfer is running
    bDone        : BOOL := FALSE; // 三段握手齐全（保持式，新循环起点清零）[-] / every handshake completed, held until a new cycle
    bFault       : BOOL := FALSE; // 故障锁存 [-] / the fault latch
    bError       : BOOL := FALSE; // 故障标志，与锁存位同源 [-] / the fault flag sharing the latch source
    iErrCode     : INT := 0;      // 错误码（锁存回放，复位沿清零）[码] / the error code replayed from the latch [code]
    ePhase       : E_DL_PltPhase := E_DL_PltPhase.eIdle; // 相位出口 [枚举] / the phase outlet [enum]
    bHoistUpCmd  : BOOL := FALSE; // 起吊命令电平 [-] / the hoist up command level
    bTraverseCmd : BOOL := FALSE; // 横移命令电平 [-] / the traverse command level
    bLowerDownCmd: BOOL := FALSE; // 下降命令电平 [-] / the lower down command level
    bSlotHold    : BOOL := FALSE; // 槽位占用等待中 [-] / waiting for the target slot
    bBeatRelease : BOOL := FALSE; // 错峰放行脉冲（单拍）[-] / the stagger release pulse, one scan wide
    nSlotActive  : INT := 0;      // 目标槽号（1 基，空闲期出 0）[号] / the target slot number, zero while idle [number]
END_VAR
VAR
    rtStart    : R_TRIG; // 启动沿，段 2 无条件刷新 / the start edge, refreshed unconditionally
    rtReset    : R_TRIG; // 复位沿，段 2 无条件刷新 / the reset edge, refreshed unconditionally
    rtSlotFree : R_TRIG; // 槽位释放沿，段 2 无条件刷新 / the slot release edge, refreshed unconditionally
    tonLift    : TON;    // 起吊超时窗，只串 eLift 相 / the hoist timeout gated by eLift
    tonTrav    : TON;    // 横移超时窗，只串 eTraverse 相 / the traverse timeout gated by eTraverse
    tonLower   : TON;    // 下降超时窗，只串 eLower 相 / the lower timeout gated by eLower
    tonSlot    : TON;    // 槽位等待超时窗，只串 eWaitSlot 相 / the slot wait timeout gated by eWaitSlot
    tonStagger : TON;    // 错峰周期窗，IN 取自身 Q 的反（自复位，FB33-2）/ the stagger period window driven by its own inverted output
    _ePhase    : E_DL_PltPhase := E_DL_PltPhase.eIdle; // 内部相位，CASE 唯一写入目标 / the internal phase, the only CASE target
    _eCause    : E_DL_PltCause := E_DL_PltCause.eNone; // 故障级成因，锁存至复位沿 / the fault cause latched until reset
    _bFault    : BOOL := FALSE; // 故障锁存位 [-] / the fault latch
    _iErrLch   : INT := 0;      // 码位锁存槽（复位沿清零）[码] / the latched code, cleared at the reset edge
    _bDone     : BOOL := FALSE; // 完成位内部锁存（清零归属：段 2 复位沿与段 3 启动沿）[-] / the internal done bit
    _bInit     : BOOL := FALSE; // 首扫初始化完成标志（R310）[-] / the first scan initialisation flag
    _bCfgOk    : BOOL := FALSE; // 时间引脚组态域内 [-] / the time pins are inside their domain
    _bSlotOk   : BOOL := FALSE; // 槽号域内 [-] / the slot number is inside its domain
    _bBeat     : BOOL := FALSE; // 本拍错峰放行（节拍脉冲与上位许可同真）[-] / the release verdict of this scan
    _bSlotEdge : BOOL := FALSE; // 槽位释放沿锁存（单拍）[-] / the one scan slot release edge
END_VAR
// 段 0｜时间量域闸与槽号越界闸：参与判据换算的引脚逐项枚举（R151）
_bCfgOk := (tLift > T#0S) AND (tTrav > T#0S) AND (tLower > T#0S) AND (tSlotWait > T#0S) AND (tStagger > T#0S); // 五个时间引脚域闸 / the five time pins domain gate
_bSlotOk := (nSlotMax >= DL_PLT_SLOT_MIN) AND (nTargetSlot >= DL_PLT_SLOT_MIN) AND (nTargetSlot <= nSlotMax); // 槽号落在 [1, nSlotMax] / the slot number inside its domain
// 段 1｜定时器与沿检测无条件周期刷新，IN 只串本相使能与锁存闸（R7、R18）
tonStagger(IN := NOT tonStagger.Q, PT := tStagger); // 错峰周期窗自复位（FB33-2，禁外部沿清零）/ the self resetting stagger window
_bBeat := tonStagger.Q AND bBeatPermit; // 本拍错峰放行判据（节拍单拍脉冲与上位许可同真）/ the release verdict of this scan
rtStart(CLK := bStart); // 启动沿无条件刷新 / unconditional refresh of the start edge
rtReset(CLK := bReset); // 复位沿无条件刷新 / unconditional refresh of the reset edge
rtSlotFree(CLK := bSlotFree); // 槽位释放沿无条件刷新 / unconditional refresh of the slot release edge
tonLift(IN := (_ePhase = E_DL_PltPhase.eLift) AND (NOT _bFault), PT := tLift); // 起吊超时窗，只串 eLift 相 / the hoist timeout gated by eLift only
tonTrav(IN := (_ePhase = E_DL_PltPhase.eTraverse) AND (NOT _bFault), PT := tTrav); // 横移超时窗，只串 eTraverse 相 / the traverse timeout gated by eTraverse only
tonLower(IN := (_ePhase = E_DL_PltPhase.eLower) AND (NOT _bFault), PT := tLower); // 下降超时窗，只串 eLower 相 / the lower timeout gated by eLower only
tonSlot(IN := (_ePhase = E_DL_PltPhase.eWaitSlot) AND (NOT _bFault), PT := tSlotWait); // 槽位超时窗，只串 eWaitSlot 相 / the slot timeout gated by eWaitSlot only
// 段 2｜首扫初始化与复位沿同块，作用域逐项声明（R310、R311）
IF (NOT _bInit) OR rtReset.Q THEN // 首扫一拍或复位沿 / the first scan or the reset edge
    _bInit := TRUE; // 首扫完成标志（复位沿重复置位同效）/ the first scan flag, the same effect on reset
    _bFault := FALSE; _eCause := E_DL_PltCause.eNone; _iErrLch := 0; // 作用域一：清锁存、清成因、清码位槽 / scope one, clear the latch, the cause and the code
    _bDone := FALSE; _ePhase := E_DL_PltPhase.eIdle; // 作用域二：清完成位并迁回空闲相 / scope two, clear the held done bit and migrate to idle
END_IF // 作用域三（单拍槽位沿 _bSlotEdge）不在此清：其每拍由启动沿段之后的沿重取行唯一写入
// 段 3｜启动沿：新循环起点同拍清完成位（R28 5.9 清零点）
IF rtStart.Q THEN _bDone := FALSE; END_IF // 完成位清零（上一循环遗留）/ clear the done bit left by the previous cycle
_bSlotEdge := rtSlotFree.Q; // 槽位释放沿重取（单拍量每拍重算，不跨拍自持）/ re-take the one scan slot release edge
// 段 4｜故障判据与锁存：未锁存才判，锁存与迁相同拍执行（R107、FB50-1④、R152）
IF NOT _bFault THEN // 未锁存才判，锁存后一律回放 / judge only while unlatched
    IF NOT _bCfgOk THEN // 时间引脚组态越域 / a time pin is out of domain
        _eCause := E_DL_PltCause.eCfgBad; _iErrLch := 301; bError := TRUE; // 故障级成因、码位与标志（R45 配对）
        _bFault := TRUE; _ePhase := E_DL_PltPhase.eFault; // 置锁存并同拍迁故障相 / latch and migrate in the same scan
    ELSIF NOT _bSlotOk THEN // 槽号越界（不起吊）/ the slot number is out of range
        _eCause := E_DL_PltCause.eSlotBad; _iErrLch := 302; bError := TRUE; // 故障级成因、码位与标志（R45 配对）
        _bFault := TRUE; _ePhase := E_DL_PltPhase.eFault; // 置锁存并同拍迁故障相 / latch and migrate in the same scan
    END_IF
END_IF
// 段 5｜相位状态机：ENUM ＋ CASE ＋ ELSE 非法相位兜底（R6、R128）
CASE _ePhase OF
E_DL_PltPhase.eIdle: // 空闲相：退出条件三（踩上节拍且目标槽已释放、目标槽未释放转等待、使能丢失则驻留）
    IF bEnable AND bStart AND _bBeat THEN // 启动电平、错峰节拍与使能同真 / the start level, the beat and the enable hold
        IF bSlotFree THEN // 目标槽已释放：直接起吊 / the target slot is free, hoist right away
            _ePhase := E_DL_PltPhase.eLift; // 迁起吊相 / migrate to the hoist phase
        ELSE // 目标槽被占：转等待相（不得起吊，互锁）/ the target slot is occupied, the interlock forbids hoisting
            _ePhase := E_DL_PltPhase.eWaitSlot; // 迁槽位等待相 / migrate to the slot wait phase
        END_IF
    END_IF
E_DL_PltPhase.eWaitSlot: // 槽位等待相：退出条件三（槽位释放沿、等待超时、使能丢失），本拍事件优先于超时（R275）
    IF NOT bEnable THEN // 使能丢失 / the enable was lost
        _ePhase := E_DL_PltPhase.eIdle; // 回空闲（命令归零由出口执行）/ back to idle, the outlet zeroes the commands
    ELSIF _bSlotEdge OR bSlotFree THEN // 槽位释放（沿或电平，电平防沿丢失）/ the slot is released either by the edge or the level
        _ePhase := E_DL_PltPhase.eLift; // 迁起吊相 / migrate to the hoist phase
    ELSIF tonSlot.Q THEN // 槽位等待超时 / the slot wait timed out
        _eCause := E_DL_PltCause.eSlotTo; _iErrLch := 306; bError := TRUE; // 故障级成因、码位与标志（R45 配对）
        _bFault := TRUE; _ePhase := E_DL_PltPhase.eFault; // 置锁存并迁故障相 / latch and migrate to the fault phase
    END_IF
E_DL_PltPhase.eLift: // 起吊相：退出条件三（起吊到位、到位超时、使能丢失）
    IF NOT bEnable THEN // 使能丢失 / the enable was lost
        _ePhase := E_DL_PltPhase.eIdle; // 回空闲 / back to idle
    ELSIF bHoistUpFb THEN // 起吊到位（拍 N 进入：本相起点、本拍行为：拒绝横移、拍 N+1 转出：横移相）
        _ePhase := E_DL_PltPhase.eTraverse; // 迁横移相 / migrate to the traverse phase
    ELSIF tonLift.Q THEN // 起吊到位超时 / the hoist limit timed out
        _eCause := E_DL_PltCause.eLiftTo; _iErrLch := 303; bError := TRUE; // 故障级成因、码位与标志（R45 配对）
        _bFault := TRUE; _ePhase := E_DL_PltPhase.eFault; // 置锁存并迁故障相 / latch and migrate to the fault phase
    END_IF
E_DL_PltPhase.eTraverse: // 横移相：退出条件三（横移到位、到位超时、使能丢失）
    IF NOT bEnable THEN // 使能丢失 / the enable was lost
        _ePhase := E_DL_PltPhase.eIdle; // 回空闲 / back to idle
    ELSIF bTravAtFb THEN // 横移到位 / the traverse limit is reached
        _ePhase := E_DL_PltPhase.eLower; // 迁下降相 / migrate to the lower phase
    ELSIF tonTrav.Q THEN // 横移到位超时 / the traverse limit timed out
        _eCause := E_DL_PltCause.eTravTo; _iErrLch := 304; bError := TRUE; // 故障级成因、码位与标志（R45 配对）
        _bFault := TRUE; _ePhase := E_DL_PltPhase.eFault; // 置锁存并迁故障相 / latch and migrate to the fault phase
    END_IF
E_DL_PltPhase.eLower: // 下降相：退出条件三（下降到位、到位超时、使能丢失）
    IF NOT bEnable THEN // 使能丢失 / the enable was lost
        _ePhase := E_DL_PltPhase.eIdle; // 回空闲 / back to idle
    ELSIF bLowerFb THEN // 下降到位（三段握手齐全）/ the lower limit is reached, all handshakes done
        _bDone := TRUE; _ePhase := E_DL_PltPhase.eDone; // 置完成位（保持至新循环起点）并迁完成相 / raise done and migrate
    ELSIF tonLower.Q THEN // 下降到位超时 / the lower limit timed out
        _eCause := E_DL_PltCause.eLowerTo; _iErrLch := 305; bError := TRUE; // 故障级成因、码位与标志（R45 配对）
        _bFault := TRUE; _ePhase := E_DL_PltPhase.eFault; // 置锁存并迁故障相 / latch and migrate to the fault phase
    END_IF
E_DL_PltPhase.eDone: // 完成相：退出条件二（启动沿消失、使能丢失）
    IF (NOT bStart) OR (NOT bEnable) THEN _ePhase := E_DL_PltPhase.eIdle; END_IF // 回空闲等下一循环 / back to idle for the next cycle
E_DL_PltPhase.eFault: // 故障相：成因锁存回放，唯一解除路径为 bReset 上升沿（R188）
    IF NOT bEnable THEN _ePhase := E_DL_PltPhase.eIdle; END_IF // 失能迁空闲（锁存位仍须复位沿解除）/ migrate to idle, the latch still needs the reset edge
ELSE // 非法相位兜底（R6、R128）/ the illegal phase fallback
    _eCause := E_DL_PltCause.ePhaseBad; _iErrLch := 307; bError := TRUE; // 故障级成因、码位与标志（R45 配对）
    _bFault := TRUE; _ePhase := E_DL_PltPhase.eFault; // 置锁存并迁故障相 / latch and migrate to the fault phase
END_CASE
IF _bFault AND (_ePhase <> E_DL_PltPhase.eFault) THEN // 段尾迁移闸：任何锁存路径不得留在业务相（FB50-1④）
    _ePhase := E_DL_PltPhase.eFault; // 统一迁故障相 / force the fault phase
END_IF
// 段 6｜统一出口：三段命令按相位单点映射，故障与失能一律归零（安全侧）
bHoistUpCmd := (_ePhase = E_DL_PltPhase.eLift) AND bEnable AND (NOT _bFault); // 起吊命令：仅起吊相且未失能未锁存 / the hoist command only in lift while enabled and unlatched
bTraverseCmd := (_ePhase = E_DL_PltPhase.eTraverse) AND bEnable AND (NOT _bFault); // 横移命令：仅横移相 / the traverse command only in traverse
bLowerDownCmd := (_ePhase = E_DL_PltPhase.eLower) AND bEnable AND (NOT _bFault); // 下降命令：仅下降相 / the lower command only in lower
bSlotHold := (_ePhase = E_DL_PltPhase.eWaitSlot) AND bEnable; // 槽位等待标志 / the slot wait flag
bBeatRelease := _bBeat AND (_ePhase = E_DL_PltPhase.eIdle) AND bEnable; // 错峰放行脉冲：单拍且仅空闲相放行 / the release pulse, one scan and idle only
nSlotActive := 0; // 空闲期槽号出零（契约：空闲不报槽号）/ report zero while idle
IF _ePhase <> E_DL_PltPhase.eIdle THEN // 非空闲期 / outside idle
    nSlotActive := nTargetSlot; // 槽号单点映射 / single point mapping of the slot number
END_IF
bBusy := bEnable AND (_ePhase <> E_DL_PltPhase.eIdle) AND (_ePhase <> E_DL_PltPhase.eDone) AND (_ePhase <> E_DL_PltPhase.eFault); // 运行位排除空闲完成与故障 / the busy bit excludes idle, done and fault
bDone := _bDone; // 完成位单点映射（保持式）/ single point mapping of the held done bit
bFault := _bFault; // 故障锁存单点映射 / single point mapping of the latch
IF _bFault THEN // 故障期回放锁存码，不在故障相按当下输入重推（R152）/ replay the latched code
    iErrCode := _iErrLch; bError := TRUE; // 锁存码回放、故障标志同源 / replay the code and share the latch source
ELSE // 非故障期 / outside fault
    iErrCode := 0; bError := FALSE; // 无故障码与无故障标志 / no code and no flag
END_IF
ePhase := _ePhase; // 相位出口单点映射 / single point mapping of the phase
END_FUNCTION_BLOCK

(* ---- FB_DL_PollAuditBank.st ---- *)
(*
  FB_DL_PollAuditBank  —  多链路轮询异常台账汇总（多实例轮询 + 首出） / Multi-link polling audit bank with first-out ledger
  分类 Category : DL_Process
  版本 Version  : 1.0.0
  来源 Source   : t1-3-oscat-network — 网络轮询审计族零检索深化
  溯源 Origin   : clean-room 实现，未复制任何源码行
  功能 Function : 1) 4 链路轮询审计：调用方轮询节拍沿 bPollTrig + 每链路当拍
                  成功量 a_bLinkOk 承载；逐链连续失败计数 auFailCnt，达 uFailTo
                  → 038E 链路异常锁存（首出链路号入 nFirstFailLink，R190 归因
                  以首出唯一承载，各链路计数独立保持）；
                  2) 恢复审计：失败计数非零链路在轮询沿收到成功 → 04B7 恢复沿
                  且计数清零；恢复不解除已锁存故障（解除仅复位沿承载）；
                  3) 故障级：038E 连续失败超阈 / 038F 组态非法（uFailTo = 0）/
                  0390 ELSE 兜底；信息级三码：首出记录 / 链路恢复 / 台账清零；
                  4) 相位机：eIdle（未使能）→ eAudit（审计中）→ eFault；
                  5) 解除式全当拍量（R240 落地），逐 BOOL 标注见段 4。
  边界 Boundary : ① 组态闸：bPollEn = FALSE 相不计数不判阈（审计仅使能相承载）；
                  ② uFailTo = 0 → 038F 锁存（连续失败阈域闸）；
                  ③ 失败计数上限钳 255（USINT 饱和前置判，防回绕）；
                  ④ 无 GVL 依赖：纯引脚输入输出，无外部变量引用，无物理 IO 地址。
  依赖 Depends  : Standard.library（R_TRIG）
  码表 Error codes（Process 段 0005，窗口 038E~0390 / 04B6~04B8）:
    16#0005_038E 故障级：链路连续失败超阈锁存（首出链路号入 nFirstFailLink），锁存至 bReset
    16#0005_038F 故障级：组态非法（失败阈 uFailTo = 0），锁存至 bReset
    16#0005_0390 故障级：相位落 ELSE 兜底，锁存至 bReset
    16#0005_04B6 信息级：首出失败记录沿（故障锁存拍）
    16#0005_04B7 信息级：链路恢复沿（失败计数非零链路收成功拍）
    16#0005_04B8 信息级：台账清零沿（复位沿清全部计数）
  修订历史 Revision :
    2026-11-19  v1.0.0  R42 首版（批次 3 · 序号 1）
*)

TYPE E_DL_PabState :
(
    eIdle   := 0,    // 未使能：不计数不判阈 / Idle, not counting
    eAudit  := 10,   // 审计中：逐链失败计数 / Audit, per-link fail counting
    eFault  := 90    // 故障：首出锁存 / Fault, latched
);
END_TYPE

FUNCTION_BLOCK FB_DL_PollAuditBank
VAR_INPUT
    a_bLinkOk    : ARRAY[0..3] OF BOOL;  // 4 链路轮询成功量（当拍量）[-] / Per-link poll success flags
    bPollTrig    : BOOL := FALSE;        // 轮询节拍沿（调用方驱动）[-] / Poll tick edge from caller
    uFailTo      : USINT := 3;           // 连续失败阈 [次]，域 > 0 / Consecutive-fail threshold
    bPollEn      : BOOL := FALSE;        // 审计使能（电平）[-] / Audit enable, level
    bReset       : BOOL := FALSE;        // 复位，上升沿清故障锁存与台账 / Reset edge clears fault and ledger
END_VAR
VAR_OUTPUT
    eState       : E_DL_PabState;     // 状态出口，段尾单点映射 / State outlet
    auFailCnt    : ARRAY[0..3] OF USINT;  // 逐链连续失败计数 [次] / Per-link consecutive-fail counts
    nFirstFailLink : DINT;            // 首出失败链路号 [0..3]，-1 = 无首出 / First failed link index
    bError       : BOOL;              // 故障锁存标志 / Fault latch flag
    nErrId       : UDINT;             // 事件码，0 = 无事件 / Event code
END_VAR
VAR
    rtPollTrig   : R_TRIG;            // 轮询节拍沿实例，无条件刷新 / Poll tick edge instance
    rtReset      : R_TRIG;            // 复位沿实例，无条件刷新 / Reset edge instance
    _eState      : E_DL_PabState := E_DL_PabState.eIdle;  // 内部相位（CASE 唯一写入目标）/ Internal phase
    _nIdx        : DINT;              // 阵列循环索引 [-] / Array loop index
    _bAllOk      : BOOL;              // 全链成功当拍量（展开式聚合）[-] / All-links-ok flag
    _nGuard      : DINT;              // WHILE/循环防死锁计数器（本件 FOR 结构性有限，仍保留计数）[-] / Loop guard counter
    _bFault      : BOOL;              // 故障锁存位（锁存量）/ Latched fault bit
    _uFault      : UDINT;             // 故障码锁存（锁存量）/ Latched fault code
    _uInfo       : UDINT;             // 信息码，每拍重算 / Transient info code
END_VAR

(* —— 段 0：沿实例无条件周期刷新（禁置于 IF/CASE 内） —— *)
_bAllOk := a_bLinkOk[0] AND a_bLinkOk[1] AND a_bLinkOk[2] AND a_bLinkOk[3];
                                        // 全链成功（当拍量，展开式聚合）
rtPollTrig(CLK := bPollTrig);           // 轮询节拍沿（每拍必调）
rtReset(CLK := bReset);                 // 复位沿（每拍必调）

(* —— 段 1：单拍量预清零（锁存量 _bFault/_uFault 与计数阵列不入清单，禁同拍抹除） —— *)
_uInfo := 16#0000_0000;             // 信息码每拍重算
nErrId := 16#0000_0000;             // 事件码缺省无事件

(* —— 段 2：复位沿 + 组态域闸（判据当拍量） —— *)
IF rtReset.Q THEN                   // rtReset.Q = 当拍量
    _bFault := FALSE;               // 清故障锁存位
    _uFault := 16#0000_0000;        // 清故障锁存码
    nFirstFailLink := -1;           // 首出链路号恢复哨兵
    FOR _nIdx := 0 TO 3 DO          // 台账逐链清零
        auFailCnt[_nIdx] := 0;      // 失败计数清零
    END_FOR
    _uInfo := 16#0005_04B8;         // 信息级：台账清零沿
END_IF
IF uFailTo = 0 THEN                 // 失败阈域闸（USINT 判等合规）
    _uFault := 16#0005_038F;        // 故障级：组态非法
    _bFault := TRUE;                // 故障标志与码位配对（R45）
END_IF

(* —— 段 3：轮询沿承载逐链审计（判据当拍量；FOR 上界 3 结构性有限，守卫计数保留） —— *)
_nGuard := 0;                       // 守卫计数预置
FOR _nIdx := 0 TO 3 DO              // 逐链审计
    _nGuard := _nGuard + 1;         // 守卫递增（FOR 结构性 ≤ 4 次，守卫仅防未来改版失控）
    IF _nGuard > 4 THEN
        EXIT;                       // 守卫兜底：异常退出（结构性不可达，防御保留）
    END_IF
    IF rtPollTrig.Q AND (_eState = E_DL_PabState.eAudit) THEN
        IF a_bLinkOk[_nIdx] THEN    // 成功：恢复审计（失败计数非零才发恢复沿）
            IF auFailCnt[_nIdx] > 0 THEN
                auFailCnt[_nIdx] := 0;              // 计数清零
                _uInfo := 16#0005_04B7;             // 信息级：链路恢复沿
            END_IF
        ELSE                        // 失败：计数递增（USINT 饱和前置判防回绕）
            IF auFailCnt[_nIdx] < 255 THEN
                auFailCnt[_nIdx] := auFailCnt[_nIdx] + 1;   // 计数递增
            END_IF
            IF (auFailCnt[_nIdx] >= uFailTo) AND (nFirstFailLink = -1) THEN
                nFirstFailLink := _nIdx;            // 首出链路号锁定（仅首个写入）
                _uFault := 16#0005_038E;            // 故障级：连续失败超阈
                _bFault := TRUE;
                _uInfo := 16#0005_04B6;             // 信息级：首出失败记录沿
            END_IF
        END_IF
    END_IF
END_FOR

(* —— 段 4：故障解除式（R240 落地，逐 BOOL 标注）：
     rtReset.Q = 当拍量；_bAllOk = 当拍量；NOT bPollEn = 当拍量。
     均不含锁存量（_bFault/_uFault），解除边真实可达（全链恢复 + 撤使能 + 复位沿）。 —— *)
IF rtReset.Q AND _bAllOk AND (NOT bPollEn) THEN
    _bFault := FALSE;               // 清故障锁存位（锁存量，仅此当拍量解除沿可清）
    _uFault := 16#0000_0000;        // 清故障锁存码（锁存量，仅本当拍量解除沿可清）
    IF _eState = E_DL_PabState.eFault THEN
        _eState := E_DL_PabState.eIdle;     // 故障相迁出：回未使能
    END_IF
END_IF

(* —— 段 5：相位机（CASE 全覆盖 + ELSE 兜底） —— *)
CASE _eState OF

E_DL_PabState.eIdle:
    IF bPollEn AND (NOT _bFault) THEN
        _eState := E_DL_PabState.eAudit;    // 使能：进审计相
    END_IF

E_DL_PabState.eAudit:
    IF (NOT _bFault) AND (NOT bPollEn) THEN
        _eState := E_DL_PabState.eIdle;     // 撤使能：回未使能相
    END_IF
    (* 首出锁存迁出在段 3 承载（置 _bFault 后段 5 次拍迁故障相） *)

E_DL_PabState.eFault:
    ;                                   // 故障相：等解除沿（段 4 承载迁出）

ELSE
    _uFault := 16#0005_0390;            // 故障级：非法相位兜底
    _bFault := TRUE;
    _eState := E_DL_PabState.eFault;    // 强制回故障相

END_CASE

(* —— 段 6：出口单点映射（名实同源；锁存码回放，禁同拍抹除） —— *)
IF _bFault THEN
    nErrId := _uFault;              // 故障锁存码回放
ELSE
    nErrId := _uInfo;               // 信息码
END_IF
bError := _bFault;                  // 故障标志与锁存位同源
eState := _eState;                  // 状态出口单点映射

END_FUNCTION_BLOCK

(* ---- FB_DL_PotlineAnodeChangeSeq.st ---- *)
// FB_DL_PotlineAnodeChangeSeq v1.0.0
// 开源溯源：clean-room 自研（族 DL_Process，ST 生态实测 0 命中，无外部代码引入）
(*
  功能: 换极十相顺控：IDLE→APPROACH→UNCLAMP→LIFT→WITHDRAW→NEWANODE→CLAMP→COVER→VERIFY→IDLE。
        联锁①LIFT 相必须 xClampOpened，违例锁存；②COVER 仅在 xClampClosed 后允许（CLAMP 后才可 COVER）；
        ③VERIFY 相阳极电流低于目标持续 30 s → 故障「新极未导通」；④FAULT 相执行器全清并锁存，仅 xReset 解除。
        fCycleS 用于相位驻留累计 _fPhaseElapsed，作 TON 之外的冗余超时判据（VERIFY 相 35 s 二次确认）。
  邻件: 与打壳机 FC_DL_PotlineCrustBreakerEnergyCalc、母线 FC_DL_PotlineBusbarShuntCalc 同族但为顺控件，不调用任何 FC。
  码表: 9321 入参非有限｜9322 组态非法(fCycleS/fCurrentTargetKA≤0)｜9323 相超时(30/10/20/30/10/60 s)
        9323 相超时（各相通用）｜9324 新极未导通｜9325 联锁违例｜9326 非法相位落 ELSE 兜底｜9327 信息级换极完成。故障码锁存至 xReset 上升沿。
  边界: 无方法块/无属性块/无全局变量/无物理 IO 地址；七 TON 单相独占且无条件刷新；xClampCmd 仅两态（TRUE 夹紧）。
*)
TYPE E_DL_AnodeChangePhase :
(
    IDLE     := 0,      // 空闲：等换极指令 [-] / Idle, waiting change command
    APPROACH := 10,     // 对位：天车移向目标槽位 [-] / Crane approaching cell
    UNCLAMP  := 20,     // 松卡具：等卡具打开反馈 [-] / Unclamping
    LIFT     := 30,     // 提极：提升残极 [-] / Lifting spent anode
    WITHDRAW := 40,     // 移出：残极移出槽位 [-] / Withdrawing anode
    NEWANODE := 50,     // 装新极：等新极就位反馈 [-] / New anode positioning
    CLAMP    := 60,     // 紧卡具：等卡具闭合反馈 [-] / Clamping
    COVER    := 70,     // 覆盖：铺保温料 [-] / Covering with crust
    VERIFY   := 80,     // 确认：新极电流导通确认 [-] / Verifying conduction
    FAULT    := 90      // 故障：锁存，仅复位沿可出 [-] / Fault latched
);
END_TYPE
FUNCTION_BLOCK FB_DL_PotlineAnodeChangeSeq
VAR_INPUT
    xEnable          : BOOL := FALSE;   // 使能，FALSE 时冻结在 IDLE [-] / Enable gate
    xStart           : BOOL := FALSE;   // 换极启动，上升沿有效 [-] / Start rising edge
    xReset           : BOOL := FALSE;   // 复位，上升沿清故障锁存 [-] / Reset rising edge
    xAtPosition      : BOOL := FALSE;   // 天车到位反馈 [-] / Crane in position
    xClampOpened     : BOOL := FALSE;   // 卡具已打开反馈 [-] / Clamp opened
    xClampClosed     : BOOL := FALSE;   // 卡具已闭合反馈 [-] / Clamp closed
    xLiftDone        : BOOL := FALSE;   // 提升完成反馈 [-] / Lift done
    xWithdrawDone    : BOOL := FALSE;   // 移出完成反馈 [-] / Withdraw done
    xNewAnodeReady   : BOOL := FALSE;   // 新极就位反馈 [-] / New anode ready
    xCoverDone       : BOOL := FALSE;   // 覆盖完成反馈 [-] / Cover done
    fAnodeCurrentKA  : REAL := 0.0;     // 实测阳极电流 [kA] / Measured anode current [kA]
    fCurrentTargetKA : REAL := 30.0;    // 目标阳极电流 [kA]，域 > 0 / Target current [kA]
    fCycleS          : REAL := 0.01;    // 任务周期 [s]，域 > 0 / Task cycle time [s]
END_VAR
VAR_OUTPUT
    ePhase       : E_DL_AnodeChangePhase;   // 相位出口，段尾单点映射 [-] / Phase outlet
    xCraneEnable : BOOL;                    // 天车使能（对位至覆盖相为真）[-] / Crane enable
    xClampCmd    : BOOL;                    // 卡具指令 TRUE 夹紧 / FALSE 松开 [-] / Clamp command
    xLiftCmd     : BOOL;                    // 提升指令（仅 LIFT 相）[-] / Lift command
    xWithdrawCmd : BOOL;                    // 移出指令（仅 WITHDRAW 相）[-] / Withdraw command
    xCoverCmd    : BOOL;                    // 覆盖指令（仅 COVER 相）[-] / Cover command
    xDone        : BOOL;                    // 换极完成单拍脉冲 [-] / Done one-shot pulse
    xFault       : BOOL;                    // 故障锁存标志 [-] / Fault latch flag
    uErrorId     : UDINT;                   // 事件码，0 = 无事件 / Event code
END_VAR
VAR
    tonApproach : TON;                      // 对位相超时 30 s，无条件刷新 / Approach timeout
    tonUnclamp  : TON;                      // 松卡具相超时 10 s，无条件刷新 / Unclamp timeout
    tonLift     : TON;                      // 提升相超时 20 s，无条件刷新 / Lift timeout
    tonWithdraw : TON;                      // 移出相超时 30 s，无条件刷新 / Withdraw timeout
    tonClamp    : TON;                      // 紧卡具相超时 10 s，无条件刷新 / Clamp timeout
    tonVerify   : TON;                      // 导通确认窗 30 s，无条件刷新 / Conduction window
    tonVerifyTo : TON;                      // 确认相总超时 60 s，无条件刷新 / Verify timeout
    tonNewAnode : TON;                      // 新极就位超时 90 s（R92 新增，防无限等待）/ New anode timeout
    tonCover    : TON;                      // 覆盖相超时 120 s（R92 新增，防铺料执行器长通）/ Cover timeout
    rtStart     : R_TRIG;                   // 启动沿实例，无条件刷新 / Start edge instance
    rtReset     : R_TRIG;                   // 复位沿实例，无条件刷新 / Reset edge instance
    _ePhase     : E_DL_AnodeChangePhase := E_DL_AnodeChangePhase.IDLE;  // 内部相位，CASE 唯一写入 / Internal phase
    _ePhasePrev : E_DL_AnodeChangePhase := E_DL_AnodeChangePhase.IDLE;  // 上拍相位快照 [-] / Previous phase snapshot
    _fElapsed   : REAL := 0.0;              // 相位驻留累计 [s]，跨周期驻留量 / Phase dwell accumulator [s]
    _xCrane     : BOOL := FALSE;            // 天车使能内部量 [-] / Internal crane enable
    _xClamp     : BOOL := FALSE;            // 卡具指令内部量 [-] / Internal clamp command
    _xLift      : BOOL := FALSE;            // 提升指令内部量 [-] / Internal lift command
    _xWithdraw  : BOOL := FALSE;            // 移出指令内部量 [-] / Internal withdraw command
    _xCover     : BOOL := FALSE;            // 覆盖指令内部量 [-] / Internal cover command
    _bFault     : BOOL := FALSE;            // 故障锁存位（锁存量，仅复位沿清）/ Latched fault bit
    _uFault     : UDINT := 16#0000;         // 故障码锁存（锁存量，仅复位沿清）/ Latched fault code
    _uInfo      : UDINT := 16#0000;         // 信息码，每拍重算 / Transient info code
END_VAR
// 段 0：定时器与沿实例无条件周期刷新（禁置于 IF/CASE 内，R7/R188）/ Unconditional refresh
rtStart(CLK := xStart);                                                     // 启动沿每拍必调 / Start edge
rtReset(CLK := xReset);                                                     // 复位沿每拍必调 / Reset edge
tonApproach(IN := (_ePhase = E_DL_AnodeChangePhase.APPROACH), PT := T#30S); // 对位超时 / Approach
tonUnclamp(IN := (_ePhase = E_DL_AnodeChangePhase.UNCLAMP), PT := T#10S);   // 松卡具超时 / Unclamp
tonLift(IN := (_ePhase = E_DL_AnodeChangePhase.LIFT), PT := T#20S);         // 提升超时 / Lift
tonWithdraw(IN := (_ePhase = E_DL_AnodeChangePhase.WITHDRAW), PT := T#30S); // 移出超时 / Withdraw
tonClamp(IN := (_ePhase = E_DL_AnodeChangePhase.CLAMP), PT := T#10S);       // 紧卡具超时 / Clamp
tonVerify(IN := (_ePhase = E_DL_AnodeChangePhase.VERIFY) AND (fAnodeCurrentKA < fCurrentTargetKA), PT := T#30S);
tonVerifyTo(IN := (_ePhase = E_DL_AnodeChangePhase.VERIFY), PT := T#60S);   // 确认相总超时 / Verify timeout
tonNewAnode(IN := (_ePhase = E_DL_AnodeChangePhase.NEWANODE), PT := T#90S);  // 新极就位超时 / New anode
tonCover(IN := (_ePhase = E_DL_AnodeChangePhase.COVER), PT := T#120S);     // 覆盖相超时 / Cover
// 段 1：单拍量与执行器量预清（锁存量 _bFault/_uFault/_fElapsed 不入清单，R187）/ One-shot clear
_uInfo := 16#0000;                  // 信息码每拍重算 / Info code recomputed
xDone := FALSE;                     // 完成脉冲缺省清 / Done pulse clear
_xCrane := FALSE;                   // 天车使能缺省关 / Crane default off
_xClamp := FALSE;                   // 卡具指令缺省松开 / Clamp default open
_xLift := FALSE;                    // 提升指令缺省关 / Lift default off
_xWithdraw := FALSE;                // 移出指令缺省关 / Withdraw default off
_xCover := FALSE;                   // 覆盖指令缺省关 / Cover default off
// 段 2：非有限闸与组态域闸（归因唯一，逐因独立码，R190）/ Gate stage
IF (fAnodeCurrentKA <> fAnodeCurrentKA) OR (fCurrentTargetKA <> fCurrentTargetKA) OR (fCycleS <> fCycleS)
   OR (ABS(fAnodeCurrentKA) >= 3.0E38) OR (ABS(fCurrentTargetKA) >= 3.0E38) OR (ABS(fCycleS) >= 3.0E38) THEN
    _uFault := 16#0002_9321;        // 故障级：入参非有限 / Fault: non-finite input
    _bFault := TRUE;                // 置故障锁存（R45 配对）/ Set fault latch
END_IF
IF (fCurrentTargetKA <= 1.0E-6) OR (fCycleS <= 1.0E-6) THEN
    _uFault := 16#0002_9322;        // 故障级：组态非法 / Fault: illegal configuration
    _bFault := TRUE;                // 置故障锁存（R45 配对）/ Set fault latch
END_IF
// 段 3：相位驻留累计（跨周期驻留量，切换拍清零）/ Phase dwell accumulation
IF _ePhase <> _ePhasePrev THEN
    _fElapsed := 0.0;               // 相位切换清零 / Reset on phase change
    _ePhasePrev := _ePhase;         // 更新快照 / Update snapshot
ELSE
    _fElapsed := _fElapsed + fCycleS;   // 同相累加周期 / Accumulate cycle
END_IF
// 段 4：复位沿（FAULT 唯一解除路径）/ Reset edge, only exit from fault
IF rtReset.Q THEN                   // rtReset.Q = 当拍量 / Reset edge per scan
    IF _ePhase = E_DL_AnodeChangePhase.FAULT THEN
        _ePhase := E_DL_AnodeChangePhase.IDLE;      // 故障相迁出回空闲 / Fault exits to idle
    END_IF
    _fElapsed := 0.0;               // 驻留累计清零（锁存量解除）/ Dwell cleared on reset
    _bFault := FALSE;               // 清故障锁存位（仅此解除沿可清）/ Clear latched bit
    _uFault := 16#0000;             // 清故障锁存码（仅此解除沿可清）/ Clear latched code
END_IF
// 段 5：相位机（本拍合法事件优先于超时，R275）/ Phase machine
CASE _ePhase OF
E_DL_AnodeChangePhase.IDLE:
    IF _bFault THEN
        _ePhase := E_DL_AnodeChangePhase.FAULT;     // 聚合故障进故障相 / Enter fault
    ELSIF rtStart.Q AND xEnable THEN
        _ePhase := E_DL_AnodeChangePhase.APPROACH;  // 启动：进对位相 / Start, approach
    END_IF
E_DL_AnodeChangePhase.APPROACH:
    _xCrane := TRUE;                                // 天车使能（同相保持）/ Crane enabled
    IF _bFault THEN
        _ePhase := E_DL_AnodeChangePhase.FAULT;     // 故障优先 / Fault first
    ELSIF NOT xEnable THEN
        _ePhase := E_DL_AnodeChangePhase.IDLE;      // 使能撤销回空闲 / Enable dropped
    ELSIF xAtPosition THEN
        _ePhase := E_DL_AnodeChangePhase.UNCLAMP;   // 到位：进松卡具相 / In position, unclamp
    ELSIF tonApproach.Q THEN
        _uFault := 16#0002_9323;                    // 故障级：对位相超时 / Approach timeout
        _bFault := TRUE;                            // 置故障锁存（R45 配对）/ Set latch
        _ePhase := E_DL_AnodeChangePhase.FAULT;     // 进故障相 / Enter fault
    END_IF
E_DL_AnodeChangePhase.UNCLAMP:
    _xCrane := TRUE;                                // 天车使能保持 / Crane enabled
    _xClamp := FALSE;                               // 卡具松开指令 / Clamp open command
    IF _bFault THEN
        _ePhase := E_DL_AnodeChangePhase.FAULT;     // 故障优先 / Fault first
    ELSIF NOT xEnable THEN
        _ePhase := E_DL_AnodeChangePhase.IDLE;      // 使能撤销回空闲（安全侧，R92 复裁补）/ Enable dropped
    ELSIF xClampOpened THEN
        _ePhase := E_DL_AnodeChangePhase.LIFT;      // 卡具已开：进提升相 / Opened, lift
    ELSIF tonUnclamp.Q THEN
        _uFault := 16#0002_9323;                    // 故障级：松卡具相超时 / Unclamp timeout
        _bFault := TRUE;                            // 置故障锁存（R45 配对）/ Set latch
        _ePhase := E_DL_AnodeChangePhase.FAULT;     // 进故障相 / Enter fault
    END_IF
E_DL_AnodeChangePhase.LIFT:
    _xCrane := TRUE;                                // 天车使能保持 / Crane enabled
    _xClamp := FALSE;                               // 卡具保持松开 / Clamp stays open
    IF _bFault THEN
        _ePhase := E_DL_AnodeChangePhase.FAULT;     // 故障优先 / Fault first
    ELSIF NOT xEnable THEN
        _ePhase := E_DL_AnodeChangePhase.IDLE;      // 使能撤销回空闲（安全侧，R92 复裁补）/ Enable dropped
    ELSIF NOT xClampOpened THEN
        _uFault := 16#0002_9325;                    // 故障级：提升时卡具未开 / Interlock violation
        _bFault := TRUE;                            // 置故障锁存（R45 配对）/ Set latch
        _ePhase := E_DL_AnodeChangePhase.FAULT;     // 进故障相 / Enter fault
    ELSIF xLiftDone THEN
        _ePhase := E_DL_AnodeChangePhase.WITHDRAW;  // 提升完成：进移出相 / Lift done, withdraw
    ELSIF tonLift.Q THEN
        _uFault := 16#0002_9323;                    // 故障级：提升相超时 / Lift timeout
        _bFault := TRUE;                            // 置故障锁存（R45 配对）/ Set latch
        _ePhase := E_DL_AnodeChangePhase.FAULT;     // 进故障相 / Enter fault
    ELSE
        _xLift := TRUE;                             // 提升指令（仅本相）/ Lift command
    END_IF
E_DL_AnodeChangePhase.WITHDRAW:
    _xCrane := TRUE;                                // 天车使能保持 / Crane enabled
    IF _bFault THEN
        _ePhase := E_DL_AnodeChangePhase.FAULT;     // 故障优先 / Fault first
    ELSIF NOT xEnable THEN
        _ePhase := E_DL_AnodeChangePhase.IDLE;      // 使能撤销回空闲（安全侧，R92 复裁补）/ Enable dropped
    ELSIF xWithdrawDone THEN
        _ePhase := E_DL_AnodeChangePhase.NEWANODE;  // 移出完成：进新极相 / Withdrawn, new anode
    ELSIF tonWithdraw.Q THEN
        _uFault := 16#0002_9323;                    // 故障级：移出相超时 / Withdraw timeout
        _bFault := TRUE;                            // 置故障锁存（R45 配对）/ Set latch
        _ePhase := E_DL_AnodeChangePhase.FAULT;     // 进故障相 / Enter fault
    ELSE
        _xWithdraw := TRUE;                         // 移出指令（仅本相）/ Withdraw command
    END_IF
E_DL_AnodeChangePhase.NEWANODE:
    _xCrane := TRUE;                                // 天车使能保持 / Crane enabled
    IF _bFault THEN
        _ePhase := E_DL_AnodeChangePhase.FAULT;     // 故障优先 / Fault first
    ELSIF NOT xEnable THEN
        _ePhase := E_DL_AnodeChangePhase.IDLE;      // 使能撤销回空闲（安全侧，R92 复裁补）/ Enable dropped
    ELSIF xNewAnodeReady THEN
        _ePhase := E_DL_AnodeChangePhase.CLAMP;     // 新极就位：进紧卡具相 / Ready, clamp
    ELSIF tonNewAnode.Q THEN
        _uFault := 16#0002_9323;                    // 故障级：相超时（新极就位，R92 复裁统一归 9323）/ Phase timeout
        _bFault := TRUE;                            // 置故障锁存 / Set latch
        _ePhase := E_DL_AnodeChangePhase.FAULT;     // 进故障相 / Enter fault
    END_IF
E_DL_AnodeChangePhase.CLAMP:
    _xCrane := TRUE;                                // 天车使能保持 / Crane enabled
    _xClamp := TRUE;                                // 卡具夹紧指令 / Clamp close command
    IF _bFault THEN
        _ePhase := E_DL_AnodeChangePhase.FAULT;     // 故障优先 / Fault first
    ELSIF NOT xEnable THEN
        _ePhase := E_DL_AnodeChangePhase.IDLE;      // 使能撤销回空闲（安全侧，R92 复裁补）/ Enable dropped
    ELSIF xClampClosed THEN
        _ePhase := E_DL_AnodeChangePhase.COVER;     // 卡具已合：进覆盖相（CLAMP 后才可 COVER）/ Go cover
    ELSIF tonClamp.Q THEN
        _uFault := 16#0002_9323;                    // 故障级：紧卡具相超时 / Clamp timeout
        _bFault := TRUE;                            // 置故障锁存（R45 配对）/ Set latch
        _ePhase := E_DL_AnodeChangePhase.FAULT;     // 进故障相 / Enter fault
    END_IF
E_DL_AnodeChangePhase.COVER:
    _xCrane := TRUE;                                // 天车使能保持 / Crane enabled
    _xClamp := TRUE;                                // 卡具保持夹紧 / Clamp stays closed
    IF _bFault THEN
        _ePhase := E_DL_AnodeChangePhase.FAULT;     // 故障优先 / Fault first
    ELSIF NOT xEnable THEN
        _ePhase := E_DL_AnodeChangePhase.IDLE;      // 使能撤销回空闲（安全侧，R92 复裁补）/ Enable dropped
    ELSIF NOT xClampClosed THEN
        _uFault := 16#0002_9325;                    // 故障级：覆盖前卡具未合 / Interlock violation
        _bFault := TRUE;                            // 置故障锁存（R45 配对）/ Set latch
        _ePhase := E_DL_AnodeChangePhase.FAULT;     // 进故障相 / Enter fault
    ELSIF xCoverDone THEN
        _ePhase := E_DL_AnodeChangePhase.VERIFY;    // 覆盖完成：进确认相 / Covered, verify
    ELSIF tonCover.Q THEN
        _uFault := 16#0002_9323;                    // 故障级：相超时（覆盖相，铺料长通，R92 复裁统一归 9323）/ Phase timeout
        _bFault := TRUE;                            // 置故障锁存 / Set latch
        _ePhase := E_DL_AnodeChangePhase.FAULT;     // 进故障相 / Enter fault
    ELSE
        _xCover := TRUE;                            // 覆盖指令（仅本相）/ Cover command
    END_IF
E_DL_AnodeChangePhase.VERIFY:
    _xClamp := TRUE;                                // 卡具保持夹紧 / Clamp stays closed
    IF _bFault THEN
        _ePhase := E_DL_AnodeChangePhase.FAULT;     // 故障优先 / Fault first
    ELSIF NOT xEnable THEN
        _ePhase := E_DL_AnodeChangePhase.IDLE;      // 使能撤销回空闲（安全侧，R92 复裁补）/ Enable dropped
    ELSIF fAnodeCurrentKA >= fCurrentTargetKA THEN
        xDone := TRUE;                              // 导通确认：完成脉冲单拍 / Conduction confirmed
        _uInfo := 16#0002_9327;                     // 信息级：换极完成 / Info: cycle done
        _ePhase := E_DL_AnodeChangePhase.IDLE;      // 回空闲 / Return to idle
    ELSIF tonVerify.Q OR (_fElapsed > 35.0) THEN
        _uFault := 16#0002_9324;                    // 故障级：新极未导通持续 30 s / Not conducting
        _bFault := TRUE;                            // 置故障锁存（R45 配对）/ Set latch
        _ePhase := E_DL_AnodeChangePhase.FAULT;     // 进故障相 / Enter fault
    ELSIF tonVerifyTo.Q THEN
        _uFault := 16#0002_9323;                    // 故障级：确认相总超时 / Verify timeout
        _bFault := TRUE;                            // 置故障锁存（R45 配对）/ Set latch
        _ePhase := E_DL_AnodeChangePhase.FAULT;     // 进故障相 / Enter fault
    END_IF
E_DL_AnodeChangePhase.FAULT:
    IF rtReset.Q THEN
        _ePhase := E_DL_AnodeChangePhase.IDLE;      // 复位沿解除（段 4 已清锁存）/ Reset releases
    END_IF
ELSE
    _uFault := 16#0002_9326;                        // 故障级：非法相位兜底（唯一占用 9326）/ Illegal phase id
    _bFault := TRUE;                                // 置故障锁存（R45 配对）/ Set latch
    _ePhase := E_DL_AnodeChangePhase.FAULT;         // 强制进故障相 / Force into fault
END_CASE
// 段 6：出口单点映射（名实双出口，R191；故障侧执行器再硬清零）/ Outlet mapping
ePhase := _ePhase;                                  // 相位出口单点映射 / Phase outlet
IF (_ePhase = E_DL_AnodeChangePhase.FAULT) OR _bFault THEN
    xCraneEnable := FALSE;                          // 故障侧天车硬零 / Fault crane hard zero
    xClampCmd := FALSE;                             // 故障侧卡具硬零 / Fault clamp hard zero
    xLiftCmd := FALSE;                              // 故障侧提升硬零 / Fault lift hard zero
    xWithdrawCmd := FALSE;                          // 故障侧移出硬零 / Fault withdraw hard zero
    xCoverCmd := FALSE;                             // 故障侧覆盖硬零 / Fault cover hard zero
    xFault := TRUE;                                 // 故障锁存回放 / Replay latched flag
    uErrorId := _uFault;                            // 故障码锁存回放 / Replay latched code
ELSE
    xCraneEnable := _xCrane;                        // 天车使能出口 / Crane enable outlet
    xClampCmd := _xClamp;                           // 卡具指令出口 / Clamp command outlet
    xLiftCmd := _xLift;                             // 提升指令出口 / Lift command outlet
    xWithdrawCmd := _xWithdraw;                     // 移出指令出口 / Withdraw command outlet
    xCoverCmd := _xCover;                           // 覆盖指令出口 / Cover command outlet
    xFault := FALSE;                                // 无故障 / No fault
    uErrorId := _uInfo;                             // 信息码每拍重算 / Transient info code
END_IF
END_FUNCTION_BLOCK

(* ---- FB_DL_PottingDispenseCtrl.st ---- *)
(*
  FB_DL_PottingDispenseCtrl  —  接线盒灌胶定量控制 / Junction-box potting dispense control
  分类 Category : DL_Process
  码位 Code     : 16#06_0_8F
  版本 Version  : 1.0.0
  溯源 Source   : LBP（Lediberg Process Library）语义借鉴 · clean-room 实现，仅借分类/参数域/命名，未复制源码
  功能 Function : 1) 称重减量法计量：灌注前后称重差折算实际灌注重量；
                  2) 双组份 A/B 混合比闭环：按设定比例分配比例输出，偏差超窗先停 A 侧（安全侧）；
                  3) 目标重量到达 + 去抖确认后置 bDoseDone（禁单拍判完成）。
  边界 Boundary : ① 称重非有限或 < 0 判 NE43 无效：冻结计量并禁止泵使能；
                  ② 混合比偏差窗上下限倒置出厂报码不运行；
                  ③ 灌注中称重回升（回流/抖动）需连续 N 拍去抖确认才判完成；
                  ④ 目标重量 <= 0 拒启动并置码；
                  ⑤ 输出三行同向：泵使能 → 比例输出 → 完成标志。
  依赖 Depends  : 无实例依赖（称重去抖自实现，避免跨件调用首拍跟踪债）

  码表 Error codes（本件子码步进 16#10，避让邻件码位）:
    16#0002_068F 故障级：组态非法（目标重量 <= 0 / 比例 <= 0 / 偏差窗倒置 / 去抖拍数 < 1）
    16#0002_069F 故障级：混合比偏差持续超窗已停 A 侧（锁存需复位）
    16#0002_06AF 信息级：称重无效计量冻结 / 目标已到去抖确认中（不置 bError）
*)

TYPE E_DL_PdcPhase :
(
    eIdle    := 0,   // 空闲待启动 / Idle
    eDose    := 10,  // 灌注计量中 / Dispensing
    eConfirm := 20,  // 目标到达去抖确认 / Target-reached debounce confirm
    eDone    := 30,  // 计量完成 / Dose done
    eFrozen  := 40,  // 称重无效冻结 / Frozen by invalid scale
    eFault   := 90   // 故障锁定 / Fault locked
);
END_TYPE

FUNCTION_BLOCK FB_DL_PottingDispenseCtrl
VAR_INPUT
    bStart        : BOOL;                           // 启动指令，上升沿生效 / Dose start, edge
    bAbort        : BOOL;                           // 中止指令，电平生效回空闲 / Abort, level
    bReset        : BOOL;                           // 复位，上升沿清故障 / Reset, clears fault
    fTargetG      : REAL := 120.0;                  // 目标灌注重量 [g]，域 > 0 / Target dose weight [g]
    fWeightAG     : REAL;                           // A 组份称重读数 [g] / Component A scale reading [g]
    fWeightBG     : REAL;                           // B 组份称重读数 [g] / Component B scale reading [g]
    fWeightStartG : REAL;                           // 灌注前称重基准 [g]（启动拍锁存）/ Pre-dose tare snapshot [g]
    fMixRatio     : REAL := 2.0;                    // A:B 混合比设定 [1]，A 份额 / Mix ratio A share [1]
    fRatioTolHi   : REAL := 10.0;                   // 比例偏差窗上限 [%]，域 > 0 / Ratio deviation window high [%]
    fRatioTolLo   : REAL := 10.0;                   // 比例偏差窗下限 [%]，域 >= 0 / Ratio deviation window low [%]
    uConfirmScans : UINT := 5;                      // 完成去抖确认拍数 [拍] / Done debounce confirm scans
    fEps          : REAL := 1.0E-6;                 // 浮点判零容差 [1] / Floating zero tolerance
END_VAR
VAR_OUTPUT
    bPumpEnable   : BOOL;                           // 计量泵使能出口 / Metering pump enable output
    fRatioOutA    : REAL;                           // A 侧比例输出 [0..1] / Component A ratio output [0..1]
    fRatioOutB    : REAL;                           // B 侧比例输出 [0..1] / Component B ratio output [0..1]
    bDoseDone     : BOOL;                           // 计量完成标志（保持型）/ Dose done flag, held
    fDosedG       : REAL;                           // 实际灌注重量 [g] = 基准 − 当前 / Actual dosed weight [g]
    bError        : BOOL;                           // 故障标志，与故障级码配对 / Fault flag
    uErrorId      : UDINT;                          // 事件码，0 = 无事件 / Event code
    eStateOut     : E_DL_PdcPhase;                  // 状态机当前态，段尾单点映射 / Phase mapped at tail
END_VAR
VAR
    _eState       : E_DL_PdcPhase := E_DL_PdcPhase.eIdle;  // 内部状态 / Internal state
    rtrStart      : R_TRIG;                         // 启动沿 / Start edge
    rtrReset      : R_TRIG;                         // 复位沿 / Reset edge
    bCfgOk        : BOOL;                           // 组态合法标志 / Configuration valid
    bScaleOkA     : BOOL;                           // A 称重本拍有效 / Scale A valid this scan
    bScaleOkB     : BOOL;                           // B 称重本拍有效 / Scale B valid this scan
    bScaleOk      : BOOL;                           // 双路称重综合有效 / Both scales valid
    fDoseAG       : REAL;                           // A 侧减量计量 [g] / A-side loss-in-weight [g]
    fDoseBG       : REAL;                           // B 侧减量计量 [g] / B-side loss-in-weight [g]
    fRatioAct     : REAL;                           // 实际混合比 [1] / Actual mix ratio [1]
    fRatioDevPct  : REAL;                           // 比例偏差 [%] / Ratio deviation [%]
    bRatioOut     : BOOL;                           // 比例超窗（电平）/ Ratio out of window
    uConfirmCnt   : UINT;                           // 完成去抖计数 [拍] / Done debounce counter
    uFault        : UDINT;                          // 锁存故障码 / Latched fault code
    uInfo         : UDINT;                          // 信息级码 / Information code
END_VAR
VAR CONSTANT
    DL_PDC_INFMAX : REAL := 1.0E30;                 // 称重有限值幅值上限 [g] / Scale finite bound [g]
END_VAR

(* === 段 0 · 实例刷新 === *)
rtrStart(CLK := bStart);                          // 每拍刷新启动沿
rtrReset(CLK := bReset);                          // 每拍刷新复位沿

(* === 段 1 · 组态闸与称重域闸 === *)
bCfgOk := (fTargetG > fEps)                       // 目标重量正域（<= 0 拒启动）
          AND (fMixRatio > fEps)                  // 比例正域
          AND (fRatioTolHi > fEps) AND (fRatioTolLo >= 0.0)   // 偏差窗不倒置且上限为正
          AND (uConfirmScans >= UINT#1)           // 去抖拍数下限
          AND (fTargetG = fTargetG) AND (fMixRatio = fMixRatio);  // NaN 自反
IF NOT bCfgOk THEN
    uFault := 16#0002_068F;                       // 故障级：组态非法
END_IF
IF rtrReset.Q AND bCfgOk THEN
    uFault := 16#0000;                            // 复位沿清锁存（解除路径可达）
END_IF
uInfo := 16#0000;                                 // 信息码每拍清零
bScaleOkA := (fWeightAG = fWeightAG) AND (fWeightAG >= 0.0) AND (fWeightAG < DL_PDC_INFMAX);  // A 路域闸
bScaleOkB := (fWeightBG = fWeightBG) AND (fWeightBG >= 0.0) AND (fWeightBG < DL_PDC_INFMAX);  // B 路域闸
bScaleOk := bScaleOkA AND bScaleOkB;              // 双路综合有效
fDosedG := 0.0;                                   // 计量值本拍重算
IF bScaleOk AND (_eState <> E_DL_PdcPhase.eIdle) THEN
    fDoseAG := fWeightStartG - fWeightAG;         // A 侧减量（基准 − 当前，回升为负）
    fDoseBG := fWeightStartG - fWeightBG;         // B 侧减量
    IF fDoseAG < 0.0 THEN
        fDoseAG := 0.0;                           // 称重回升不外推负计量（去抖确认承担）
    END_IF
    IF fDoseBG < 0.0 THEN
        fDoseBG := 0.0;                           // 同上 B 侧
    END_IF
    fDosedG := fDoseAG + fDoseBG;                 // 实际灌注 = 双侧减量和
END_IF

(* === 段 2 · 混合比闭环判据（本拍重算）=== *)
fRatioAct := 1.0;                                 // 实际比缺省 1（防除零哨兵）
fRatioDevPct := 0.0;                              // 偏差缺省 0
bRatioOut := FALSE;                               // 超窗标志本拍重算
IF bScaleOk AND (fDoseBG > fEps) THEN
    fRatioAct := fDoseAG / fDoseBG;               // A/B 实际比（分母已判零）
    fRatioDevPct := ABS(fRatioAct - fMixRatio) / fMixRatio * 100.0;   // 相对偏差 [%]（分母组态闸已保证 > 0）
    bRatioOut := (fRatioDevPct > fRatioTolHi + fEps) OR (fRatioDevPct < -fRatioTolLo - fEps);  // 超窗判定
END_IF

(* === 段 3 · 主状态机（ENUM + CASE，含 ELSE 兜底）=== *)
CASE _eState OF
E_DL_PdcPhase.eIdle :
    bPumpEnable := FALSE;                         // 空闲泵停
    fRatioOutA := 0.0;                            // 比例输出清零
    fRatioOutB := 0.0;
    IF uFault <> 16#0000 THEN
        _eState := E_DL_PdcPhase.eFault;          // 故障优先
    ELSIF NOT bScaleOk THEN
        _eState := E_DL_PdcPhase.eFrozen;         // 称重无效进冻结
    ELSIF rtrStart.Q AND bCfgOk THEN
        _eState := E_DL_PdcPhase.eDose;           // 启动沿进灌注相
    END_IF

E_DL_PdcPhase.eDose :
    bPumpEnable := bScaleOk AND (uFault = 16#0000);   // 称重无效/故障即停泵（安全侧）
    fRatioOutA := fMixRatio / (fMixRatio + 1.0);  // A 份额按设定比分配（分母 > 0 组态闸保证）
    fRatioOutB := 1.0 - fRatioOutA;               // B 份额互补
    IF bRatioOut THEN
        fRatioOutA := 0.0;                        // 比例超窗先停 A 侧（安全侧）
        uFault := 16#0002_069F;                   // 故障级：混合比偏差持续超窗停 A 侧（锁存）
        _eState := E_DL_PdcPhase.eFault;          // 转故障相
    ELSIF NOT bScaleOk THEN
        uInfo := 16#0002_06AF;                    // 信息级：称重无效计量冻结
        _eState := E_DL_PdcPhase.eFrozen;         // 转冻结相
    ELSIF bAbort THEN
        _eState := E_DL_PdcPhase.eIdle;           // 中止回空闲
    ELSIF fDosedG >= fTargetG THEN
        uInfo := 16#0002_06AF;                    // 信息级：目标已到去抖确认中
        uConfirmCnt := UINT#0;                    // 确认计数从 0 起算
        _eState := E_DL_PdcPhase.eConfirm;        // 进确认相（禁单拍判完成）
    END_IF

E_DL_PdcPhase.eConfirm :
    bPumpEnable := FALSE;                         // 确认相泵已停（目标到即停）
    IF bScaleOk AND (fDosedG >= fTargetG - fEps) THEN
        uConfirmCnt := uConfirmCnt + UINT#1;      // 稳定保持计数累加
        IF uConfirmCnt >= uConfirmScans THEN
            bDoseDone := TRUE;                    // 连续 N 拍稳定在目标域：完成
            _eState := E_DL_PdcPhase.eDone;       // 转完成相
        END_IF
    ELSE
        uConfirmCnt := UINT#0;                    // 回落：计数清零重计
        IF bScaleOk THEN
            _eState := E_DL_PdcPhase.eDose;       // 未达稳态回灌注相（欠量补灌）
        ELSE
            _eState := E_DL_PdcPhase.eFrozen;     // 称重丢失转冻结
        END_IF
    END_IF

E_DL_PdcPhase.eDone :
    bPumpEnable := FALSE;                         // 完成相泵停
    bDoseDone := TRUE;                            // 完成保持（防同拍抹除）
    IF rtrStart.Q AND bScaleOk THEN
        bDoseDone := FALSE;                       // 新启动沿重开计量
        _eState := E_DL_PdcPhase.eDose;           // 回灌注相
    ELSIF NOT bScaleOk THEN
        _eState := E_DL_PdcPhase.eFrozen;         // 称重丢失转冻结（完成标志保持）
    END_IF

E_DL_PdcPhase.eFrozen :
    bPumpEnable := FALSE;                         // 冻结相禁泵使能（计量冻结）
    IF bScaleOk AND (uFault = 16#0000) THEN
        _eState := E_DL_PdcPhase.eDose;           // 称重恢复回灌注（解除路径可达，欠量续灌）
    END_IF

E_DL_PdcPhase.eFault :
    bPumpEnable := FALSE;                         // 故障相禁泵
    IF uFault = 16#0000 THEN
        _eState := E_DL_PdcPhase.eIdle;           // 解锁回空闲
    END_IF

ELSE
    _eState := E_DL_PdcPhase.eFault;              // 非法状态拦截
    uFault := 16#0002_068F;                       // 故障级：相 ID 越界复用组态码段
END_CASE

(* === 段 4 · 输出映射 === *)
bError := (uFault <> 16#0000);                    // 故障标志仅由故障级码置位（R45 配对）
IF bError THEN
    uErrorId := uFault;                           // 故障级优先上报
ELSE
    uErrorId := uInfo;                            // 否则上报信息级码
END_IF
eStateOut := _eState;                             // 输出枚举段尾单点映射（N2 规则）
END_FUNCTION_BLOCK

(* ---- FB_DL_PouchVacuumSeal.st ---- *)
(*
  FB_DL_PouchVacuumSeal  —  铝塑膜真空封装顺控（真空度窗 + 封头温度 + 封合延时） / Aluminium-laminate pouch vacuum sealing with vacuum window, head-temperature window and seal dwell
  分类 Category : DL_Process
  版本 Version  : 1.0.0
  来源 Source   : roadmap-li-p1 — 锂电软包封装工站真缺口
  溯源 Origin   : 道莅 clean-room 实现；真空封装「抽真空-封合-冷却」时序与真空度/温度窗判据为公开工艺逻辑，未复制任何源码行
  功能 Function : 1) 三段顺控：eEvac 抽真空（真空度 fVacKpa 达 fVacTargetKpa 容差带内）→
                  eSeal 封合（封头温度在 [fSealTempLoC, fSealTempHiC] 窗内且 tSeal 到时）→
                  eCool 冷却（tCool 到时）→ eDone；2) 抽真空超时 tEvacTmo 保护；
                  3) 封合相温度越窗即故障，温度窗判据为双向容差式；
                  4) 故障级单码 039E，归因由 eCause 独立成员承载（R190）；
                  5) 信息级 04C6 = 封装循环完成沿；6) 解除式全当拍量（R240）。
  接口 Interface: 输入真空度/封头温度/三个时间量/命令位；输出状态/真空镜像/窗内镜像/原因/码
  边界 Boundary : ① 组态闸：fVacTargetKpa > 0.0（目标真空度按正压差量纲给出，域 > 0）、
                  fSealTempHiC <= fSealTempLoC、三个时间量 <= T#0S → 039E 锁存；
                  ② 真空度判据用 fVacKpa - fVacTargetKpa 的容差带（|Δ| <= fVacTolKpa），
                  禁用 = / <> 判等；③ 封头温度判据同样容差式；
                  ④ 三个 TON + 一个 R_TRIG 全部段 0 无条件每周期调用，IN 由相位派生，
                  相切换自动复位 ET；⑤ 故障相迁出唯一路径 = bReset 上升沿；
                  ⑥ 零全局耦合：无 GVL / VAR_EXTERNAL / %I %Q %M。
  依赖 Depends  : Standard.library（TON / R_TRIG）
  码表 Error codes（Process 段 0005，故障窗口 039E / 信息窗口 04C6）:
    16#0005_039E 故障级：真空封装故障总码（组态非法 / 抽真空超时 / 封头温度越窗），
                 锁存至 bReset 上升沿；逐成因归因见 eCause，不新增码位（派单硬约束单码）
    16#0005_04C6 信息级：封装循环完成沿（冷却完成进 eDone 单拍）
  修订历史 Revision :
    2026-11-19  v1.0.0  R43 首版（批次 1 · 序号 2）
*)

TYPE E_DL_PvsState :
(
    eIdle   := 0,     // 未使能待启动 / Idle, waiting start
    eEvac   := 10,    // 抽真空中 / Evacuating
    eSeal   := 20,    // 封合中（温度窗 + 延时） / Sealing under temperature window
    eCool   := 30,    // 冷却中 / Cooling
    eDone   := 50,    // 循环完成 / Done
    eFault  := 90     // 故障锁存相 / Fault latched phase
);
END_TYPE

TYPE E_DL_PvsCause :
(
    eNone       := 0,    // 无故障成因 / No cause
    eCfgIllegal := 1,    // 组态非法 / Illegal configuration
    eEvacTmo    := 2,    // 抽真空超时 / Evacuation timeout
    eSealTemp   := 3     // 封头温度越窗 / Seal head temperature out of window
);
END_TYPE

FUNCTION_BLOCK FB_DL_PouchVacuumSeal
VAR_INPUT
    fVacKpa      : REAL := 0.0;        // 实测真空度 [kPa]，相对大气压正压差量纲 / Measured vacuum level
    fVacTargetKpa: REAL := 95.0;       // 目标真空度 [kPa]，域 > 0 / Target vacuum level
    fVacTolKpa   : REAL := 2.0;        // 真空度容差带 [kPa]，域 > 0 / Vacuum tolerance band
    fSealTempC   : REAL := 0.0;        // 实测封头温度 [°C] / Measured seal head temperature
    fSealTempLoC : REAL := 150.0;      // 封头温度窗下限 [°C] / Head temperature low limit
    fSealTempHiC : REAL := 175.0;      // 封头温度窗上限 [°C] / Head temperature high limit
    tEvacTmo     : TIME := T#20S;      // 抽真空超时 [ms]，域 > 0 / Evacuation timeout
    tSeal        : TIME := T#3S;       // 封合延时 [ms]，域 > 0 / Seal dwell
    tCool        : TIME := T#2S;       // 冷却时长 [ms]，域 > 0 / Cooling duration
    bStart       : BOOL := FALSE;      // 启动命令（电平）[-] / Start command
    bReset       : BOOL := FALSE;      // 复位命令，上升沿清故障 [-] / Reset edge
END_VAR
VAR_OUTPUT
    eState       : E_DL_PvsState;      // 状态出口，段 6 单点映射 / State outlet
    eCause       : E_DL_PvsCause;      // 故障成因出口（R190） / Fault cause outlet
    fVacKpaOut   : REAL;               // 真空度镜像 [kPa] / Vacuum mirror
    bVacOk       : BOOL;               // 真空度达窗镜像 [-] / Vacuum reached mirror
    bTempOk      : BOOL;               // 封头温度在窗镜像 [-] / Head temperature in window
    bCycleDone   : BOOL;               // 循环完成标志 [-] / Cycle done flag
    bError       : BOOL;               // 故障锁存标志 [-] / Fault latch flag
    nErrId       : UDINT;              // 事件码，0 = 无事件 / Event code
END_VAR
VAR
    _eState      : E_DL_PvsState := E_DL_PvsState.eIdle;   // 内部相位（CASE 唯一写入目标） / Internal phase
    _eCause      : E_DL_PvsCause := E_DL_PvsCause.eNone;   // 故障成因锁存（锁存量） / Latched cause
    tonEvac      : TON;                // 抽真空超时实例，每周期无条件调用 / Evacuation timeout timer
    tonSeal      : TON;                // 封合延时实例，每周期无条件调用 / Seal dwell timer
    tonCool      : TON;                // 冷却计时实例，每周期无条件调用 / Cooling timer
    rtReset      : R_TRIG;             // 复位沿实例，每周期无条件调用 / Reset edge
    _bVacOk      : BOOL;               // 真空度达窗当拍量 [-] / Vacuum window verdict
    _bTempOk     : BOOL;               // 温度在窗当拍量 [-] / Temperature window verdict
    _bCfgBad     : BOOL;               // 组态非法当拍量 [-] / Config illegal
    _bFault      : BOOL;               // 故障锁存位（锁存量） / Latched fault bit
    _uFault      : UDINT;              // 故障码锁存（锁存量） / Latched fault code
    _uInfo       : UDINT;              // 信息码，每拍重算 / Transient info code
END_VAR

(* —— 段 0：沿实例与定时器无条件周期刷新 —— *)
_bVacOk := ABS(fVacKpa - fVacTargetKpa) <= fVacTolKpa;                          // 真空度容差窗判据 / Vacuum tolerance window verdict
_bTempOk := (fSealTempC >= fSealTempLoC - 1.0E-6) AND (fSealTempC <= fSealTempHiC + 1.0E-6);  // 温度容差窗判据 / Temperature window verdict
_bCfgBad := (fVacTargetKpa <= 0.0) OR (fVacTolKpa <= 0.0)
            OR (fSealTempHiC <= fSealTempLoC) OR (tEvacTmo <= T#0S)
            OR (tSeal <= T#0S) OR (tCool <= T#0S);                              // 组态非法当拍量 / Config illegal, current scan
rtReset(CLK := bReset);                                                        // 复位沿，每拍必调 / Reset edge refresh
tonEvac(IN := (_eState = E_DL_PvsState.eEvac), PT := tEvacTmo);                // 抽真空超时计时  / Evacuation timer
tonSeal(IN := (_eState = E_DL_PvsState.eSeal), PT := tSeal);                   // 封合延时计时 / Seal dwell timer
tonCool(IN := (_eState = E_DL_PvsState.eCool), PT := tCool);                   // 冷却计时 / Cooling timer

(* —— 段 1：单拍量预清零（锁存量不入清单，禁同拍抹除 R187） —— *)
_uInfo := 16#0000_0000;            // 信息码每拍重算 / Info recomputed
fVacKpaOut := 0.0;                 // 真空镜像缺省 0 / Vacuum mirror default
bVacOk := FALSE;                   // 达窗镜像缺省 FALSE / Vacuum flag default
bTempOk := FALSE;                  // 温度镜像缺省 FALSE / Temperature flag default
bCycleDone := FALSE;               // 完成标志缺省 FALSE / Done default
nErrId := 16#0000_0000;            // 事件码缺省无事件 / Event code default

(* —— 段 2：复位沿 + 组态域闸（当拍量判据） —— *)
IF rtReset.Q THEN                              // rtReset.Q = 当拍量 / current scan
    _bFault := FALSE;                          // 清故障锁存位（锁存量） / Clear fault latch
    _uFault := 16#0000_0000;                   // 清故障锁存码（锁存量） / Clear fault code
    _eCause := E_DL_PvsCause.eNone;            // 清成因（锁存量） / Clear cause
    IF _eState = E_DL_PvsState.eFault THEN
        _eState := E_DL_PvsState.eIdle;        // 故障相迁出：回未使能 / Fault exit to idle
    END_IF
END_IF
IF _bCfgBad THEN                               // 组态域闸 / Config gate
    _uFault := 16#0005_039E;                   // 故障级：真空封装故障总码 / Process fault code
    _eCause := E_DL_PvsCause.eCfgIllegal;      // 归因：组态非法 / Cause: illegal config
    _bFault := TRUE;                           // 标志与码位配对（R45） / Flag paired with code
END_IF

(* —— 段 3：抽真空超时与封合温度越窗（判据当拍量） —— *)
IF (NOT _bFault) AND tonEvac.Q THEN            // 抽真空超时 / Evacuation timeout
    _uFault := 16#0005_039E;                   // 故障级：总码 / Public code
    _eCause := E_DL_PvsCause.eEvacTmo;         // 归因：抽真空超时 / Cause: evac timeout
    _bFault := TRUE;
END_IF
IF (NOT _bFault) AND (_eState = E_DL_PvsState.eSeal) AND (NOT _bTempOk) THEN  // 封合期温度越窗 / Seal temp deviation
    _uFault := 16#0005_039E;
    _eCause := E_DL_PvsCause.eSealTemp;        // 归因：封头温度越窗 / Cause: seal temperature
    _bFault := TRUE;
END_IF

(* —— 段 4：故障解除式（R240；全当拍量）：rtReset.Q / NOT _bCfgBad / NOT tonEvac.Q / NOT tonSeal.Q 皆当拍量 —— *)
IF rtReset.Q AND (NOT _bCfgBad) AND (NOT tonEvac.Q) AND (NOT tonSeal.Q) THEN
    _bFault := FALSE;                          // 清故障锁存位（锁存量） / Clear fault latch
    _uFault := 16#0000_0000;                   // 清故障锁存码（锁存量） / Clear fault code
    _eCause := E_DL_PvsCause.eNone;            // 清成因（锁存量） / Clear cause
END_IF

(* —— 段 4A：故障锁存相位迁移闸 —— *)
IF _bFault AND (_eState <> E_DL_PvsState.eFault) THEN
    _eState := E_DL_PvsState.eFault;           // 锁存即入故障相 / Latch enters fault phase
END_IF

(* —— 段 5：相位机（CASE 全覆盖 + ELSE 兜底） —— *)
CASE _eState OF

E_DL_PvsState.eIdle:
    IF bStart AND (NOT _bFault) THEN           // 启动条件 / Start gate
        _eState := E_DL_PvsState.eEvac;        // 进抽真空相 / Enter evacuation
    END_IF

E_DL_PvsState.eEvac:
    IF _bVacOk THEN                            // 出口 1：真空度达窗 / Vacuum reached
        _eState := E_DL_PvsState.eSeal;        // 进封合相 / Enter sealing
    ELSIF NOT bStart THEN                      // 出口 2：撤启动（R98 双出口） / Start released
        _eState := E_DL_PvsState.eIdle;
    END_IF

E_DL_PvsState.eSeal:
    IF tonSeal.Q AND _bTempOk THEN             // 封合延时到且温度在窗 / Dwell done within window
        _eState := E_DL_PvsState.eCool;        // 进冷却相 / Enter cooling
    ELSIF NOT bStart THEN                      // 撤启动：中止 / Abort
        _eState := E_DL_PvsState.eIdle;
    END_IF

E_DL_PvsState.eCool:
    IF tonCool.Q THEN                          // 冷却到时 / Cooling elapsed
        _uInfo := 16#0005_04C6;                // 信息级：循环完成沿 / Info: cycle complete edge
        _eState := E_DL_PvsState.eDone;        // 进完成相 / Enter done
    ELSIF NOT bStart THEN                      // 撤启动：中止 / Abort
        _eState := E_DL_PvsState.eIdle;
    END_IF

E_DL_PvsState.eDone:
    IF NOT bStart THEN                         // 撤启动回空闲 / Start released returns idle
        _eState := E_DL_PvsState.eIdle;
    END_IF

E_DL_PvsState.eFault:
    ;                                          // 故障相：仅段 4 复位沿可迁出 / Only reset exits

ELSE
    _uFault := 16#0005_039E;                   // 故障级：非法相位兜底（归并总码） / Illegal phase fallback
    _eCause := E_DL_PvsCause.eCfgIllegal;      // 归因：相位非法归并组态 / Cause: phase illegal
    _bFault := TRUE;
    _eState := E_DL_PvsState.eFault;           // 强制回故障相 / Force fault phase

END_CASE

(* —— 段 6：出口单点映射（名实同源；锁存码回放） —— *)
fVacKpaOut := fVacKpa;                         // 真空镜像 / Vacuum mirror
bVacOk := _bVacOk AND (NOT _bFault);           // 达窗镜像 / Vacuum verdict mirror
bTempOk := _bTempOk AND (NOT _bFault);         // 温度窗镜像 / Temperature verdict mirror
bCycleDone := (_eState = E_DL_PvsState.eDone);// 完成标志 / Done flag
IF _bFault THEN
    nErrId := _uFault;                         // 故障锁存码回放 / Replay latched code
ELSE
    nErrId := _uInfo;                          // 信息码 / Transient info
END_IF
bError := _bFault;                             // 故障标志同源 / Flag from latch
eState := _eState;                             // 状态出口 / State outlet
eCause := _eCause;                             // 成因出口 / Cause outlet

END_FUNCTION_BLOCK
